      $ 2057 "Vial_liq_pick_3" "breakAfter"
      movel(Vial_liq_pick_3_p, a=0.5, v=0.1)
      $ 2058 "Vial_liq_pick_4" "breakAfter"
      movel(Vial_liq_pick_4_p, a=0.5, v=0.1)
      # begin: URCap Program Node
      #   Source: Robotiq_Grippers, 3.17.0.105337, Robotiq Inc.
      #   Type: Gripper
      $ 2059 "Gripper Close (1)"
      if not(gripper_connected[0]):
        popup("Gripper 1 must be connected to run this program.", "No connection", False, True, True)
      end
      if not(rq_is_gripper_activated("1")):
        popup("Gripper 1 is not activated. Go to Installation tab > Gripper to activate it and run the program again.", "Not activated", False, True, True)
      end
      rq_set_pos_spd_for(255, 82, 71, "1")
      rq_wait_pos_spe_for_request(255, 82, 71, "1")
      rq_go_to("1")
      rq_wait("1")
      # end: URCap Program Node
      $ 2060 "Wait: 1.0"
      sleep(1.0)
      $ 2061 "Set GRP_3F_Open=On"
      set_standard_digital_out(5, True)
      $ 2062 "Wait: 0.5"
      sleep(0.5)
      $ 2063 "Vial_liq_abov_2" "breakAfter"
      movel(Vial_liq_abov_2_p, a=0.3, v=0.05, r=0.05)
      $ 2064 "MoveL"
      $ 2065 "Liquid_midway_1" "breakAfter"
      movel(Liquid_midway_1_p, a=0.5, v=0.1)
      $ 2066 "Loop 3 times"
      Loop_1 = 0
      while (Loop_1 < 3):
        $ 2067 "shake_3" "breakAfter"
        movel(shake_3_p, a=2.0, v=0.5)
        $ 2068 "shake_4" "breakAfter"
        movel(shake_4_p, a=2.0, v=0.5)
        Loop_1 = Loop_1 + 1
      end
      $ 2069 "drop_above_3" "breakAfter"
      movel(drop_above_3_p, a=0.5, v=0.1)
      $ 2070 "drop_above_4" "breakAfter"
      movel(drop_above_4_p, a=0.5, v=0.1)
      $ 2071 "liq_tran_3" "breakAfter"
      movel(liq_tran_3_p, a=0.5, v=0.05, r=0.008)
      $ 2072 "Wait: 1.0"
      sleep(1.0)
      $ 2073 "drop_above_5" "breakAfter"
      movel(drop_above_5_p, a=0.5, v=0.1)
      $ 2074 "Waypoint_92" "breakAfter"
      movel(Waypoint_92_p, a=0.5, v=0.1)
      $ 2075 "liq_tran_4" "breakAfter"
      movel(liq_tran_4_p, a=0.5, v=0.05)
      $ 2076 "Wait: 1.0"
      sleep(1.0)
      $ 2077 "drop_above_6" "breakAfter"
      movel(drop_above_6_p, a=0.5, v=0.1)
      $ 2078 "drop_above_7" "breakAfter"
      movel(drop_above_7_p, a=0.5, v=0.1)
      $ 2079 "Liquid_midway_2" "breakAfter"
      movel(Liquid_midway_2_p, a=0.5, v=0.1)
      $ 2080 "MoveL"
      $ 2081 "Vial_drop_abo_1" "breakAfter"
      movel(Vial_drop_abo_1_p, a=0.5, v=0.1)
      $ 2082 "Vial_liq_drop_1" "breakAfter"
      movel(Vial_liq_drop_1_p, a=0.5, v=0.1)
      # begin: URCap Program Node
      #   Source: Robotiq_Grippers, 3.17.0.105337, Robotiq Inc.
      #   Type: Gripper
      $ 2083 "Gripper Open (1)"
      if not(gripper_connected[0]):
        popup("Gripper 1 must be connected to run this program.", "No connection", False, True, True)
      end
      if not(rq_is_gripper_activated("1")):
        popup("Gripper 1 is not activated. Go to Installation tab > Gripper to activate it and run the program again.", "Not activated", False, True, True)
      end
      rq_set_pos_spd_for(0, 82, 71, "1")
      rq_wait_pos_spe_for_request(0, 82, 71, "1")
      rq_go_to("1")
      rq_wait("1")
      # end: URCap Program Node
      $ 2084 "Vial_drop_abo_2" "breakAfter"
      movel(Vial_drop_abo_2_p, a=0.5, v=0.1)
    elif (34 == switch_1):
      $ 2085 "Case 34"
      $ 2086 "Task≔'Dosing'"
      global Task="Dosing"
      $ 2087 "tilt_to_home()"
      tilt_to_home()
      $ 2088 "Powder dosing all"
      $ 2089 "tilt_angle_sent≔0.0"
      global tilt_angle_sent=0.0
      $ 2090 "send_target_info()"
      send_target_info()
      $ 2092 "prev_spat≔''"
      global prev_spat=""
      $ 2093 "spatula≔''"
      global spatula=""
      $ 2094 "scoop_status≔'normal'"
      global scoop_status="normal"
      $ 2095 "send_powder_info()"
      send_powder_info()
      $ 2096 "Set AO[0]=0.0"
      set_standard_analog_out(0, 0.0)
      $ 2097 "Wait: 0.2"
      sleep(0.2)
      $ 2098 "reach pots decapping pose"
      # begin: URCap Program Node
      #   Source: SensoPart VISOR Robotic, 2.0.6, SensoPart Industriesensorik GmbH
      #   Type: VISOR Robotic App
      $ 2104 "VISOR Easy Pick"
      def visorFuncEasyPick_14c2cb():
        # begin: URCap Program Node
        #   Source: SensoPart VISOR Robotic, 2.0.6, SensoPart Industriesensorik GmbH
        #   Type: Easy Pick Setup
        $ 2105 "# 1 Setup" "noBreak"
        local easyPickVisorId = 1
        local easyPickArmMounted = True
        local easyPickSetJob = True
        local easyPickJobName = "Weight_scale"
        local easyPickAtImgAcq = False
        local easyPickImgAcqPose = Trigger
        # end: URCap Program Node
        # begin: URCap Program Node
        #   Source: SensoPart VISOR Robotic, 2.0.6, SensoPart Industriesensorik GmbH
        #   Type: Process
        $ 2106 "Process" "noBreak"
        local easyPickObjTaken = False
        local easyPickTrigger = False
        local easyPickPoseIdx = 0
        local easyPickPose = p[0,0,0,0,0,0]
        def easyPickFuncTrigger(visorId, setJob, jobName, arm):
        if (setJob):
          visor_changeJob(visorId, jobName, 6000)
        end
        if (arm):
          visor_trigger(visorId, 6000, "arm")
        else:
          visor_trigger(visorId, 6000)
        end
        global easyPickParts_4=visor_partsFound(visorId)
        visor_easyPickUpdate(visorId, "parts", visor_partsFound(visorId))
        return visor_getPose3d(visorId, 0)
      end
      while (not easyPickObjTaken):
        easyPickTrigger = (easyPickCount_4 >= visor_partsFound(easyPickVisorId)) or (easyPickCount_4 > 9) or (not visor_easyPickCheckIdent("850a49", easyPickVisorId))
        if (easyPickTrigger):
          easyPickCount_4 = 0
        end
        easyPickPoseIdx = easyPickCount_4
        easyPickPose = visor_getPose3d(easyPickVisorId, easyPickPoseIdx)
        visor_easyPickUpdate(easyPickVisorId, "counter", easyPickPoseIdx)
        # begin: URCap Program Node
        #   Source: SensoPart VISOR Robotic, 2.0.6, SensoPart Industriesensorik GmbH
        #   Type: Image Acquisition Pose
        $ 2107 "Image Acquisition Pose" "noBreak"
        if (easyPickTrigger):
          if (not easyPickAtImgAcq):
            movej(pose_trans(easyPickImgAcqPose,p[0.0000,0.0000,-0.0000,0.0000,0.0000,0.0000]),a=1.3963,v=1.0472,t=0.000000,r=0.000000)
            easyPickAtImgAcq = True
          end
          easyPickPose = easyPickFuncTrigger(easyPickVisorId, easyPickSetJob, easyPickJobName, easyPickArmMounted)
        end
        # end: URCap Program Node
        # begin: URCap Program Node
        #   Source: SensoPart VISOR Robotic, 2.0.6, SensoPart Industriesensorik GmbH
        #   Type: Object Detected
        $ 2108 "Object Detected" "noBreak"
        if (visor_partsFound(easyPickVisorId) > 0):
          $ 2109 "Open Gripper" "noBreak"
          $ 2110 "weight_value≔get_weight()" "noBreak"
          global weight_value=get_weight()
          $ 2111 "Wait: 0.5" "noBreak"
          sleep(0.5)
          $ 2112 "diff≔target_weight-weight_value" "noBreak"
          global diff=target_weight-weight_value
          $ 2113 "compute_level_percent(W_now, weight_value)" "noBreak"
          compute_level_percent(W_now, weight_value)
          $ 2114 "send_level_info()" "noBreak"
          send_level_info()
          $ 2115 "spatula≔select_spatula(Flowability, level, diff, bulk_density, mouth_d)" "noBreak"
          global spatula=select_spatula(Flowability, level, diff, bulk_density, mouth_d)
          $ 2116 "Wait: 0.2" "noBreak"
          sleep(0.2)
          $ 2117 "send_spatula_info()" "noBreak"
          send_spatula_info()
          $ 2118 "Pick spatula" "noBreak"
          $ 2119 "If spatula ≟ 'spatula_L'" "noBreak"
          if (spatula  ==  "spatula_L"):
            $ 2120 "MoveJ" "noBreak"
            $ 2121 "Spatula_otw" "noBreak"
            movej(get_inverse_kin(Spatula_otw_p, qnear=Spatula_otw_q), a=1.3962634015954636, v=1.0471975511965976)
            $ 2122 "pick_spat_L_abv" "noBreak"
            movej(get_inverse_kin(pick_spat_L_abv_p, qnear=pick_spat_L_abv_q), a=1.3962634015954636, v=1.0471975511965976)
            $ 2123 "MoveL" "noBreak"
            $ 2124 "spat_L_pick" "noBreak"
            movel(spat_L_pick_p, a=1.2, v=0.25)
            # begin: URCap Program Node
            #   Source: Robotiq_Grippers, 3.17.0.105337, Robotiq Inc.
            #   Type: Gripper
            $ 2125 "Gripper Close (1)" "noBreak"
            if not(gripper_connected[0]):
              popup("Gripper 1 must be connected to run this program.", "No connection", False, True, True)
            end
            if not(rq_is_gripper_activated("1")):
              popup("Gripper 1 is not activated. Go to Installation tab > Gripper to activate it and run the program again.", "Not activated", False, True, True)
            end
            rq_set_pos_spd_for(255, 0, 77, "1")
            rq_wait_pos_spe_for_request(255, 0, 77, "1")
            rq_go_to("1")
            rq_wait("1")
            # end: URCap Program Node
            $ 2126 "spat_L_lift" "noBreak"
            movel(spat_L_lift_p, a=1.2, v=0.25, r=0.01)
            $ 2127 "spat_L_side" "noBreak"
            movel(spat_L_side_p, a=1.2, v=0.25, r=0.01)
            $ 2128 "spat_L_up" "noBreak"
            movel(spat_L_up_p, a=1.2, v=0.25, r=0.05)
            $ 2129 "MoveJ" "noBreak"
            $ 2130 "Spatula_otw" "noBreak"
            movej(get_inverse_kin(Spatula_otw_p, qnear=Spatula_otw_q), a=1.3962634015954636, v=1.0471975511965976)
          else:
            $ 2131 "ElseIf spatula ≟'spatula_M'" "noBreak"
            if (spatula  == "spatula_M"):
              $ 2132 "MoveJ" "noBreak"
              $ 2133 "Spatula_otw" "noBreak"
              movej(get_inverse_kin(Spatula_otw_p, qnear=Spatula_otw_q), a=1.3962634015954636, v=1.0471975511965976)
              $ 2134 "spat_M_up" "noBreak"
              movej(get_inverse_kin(spat_M_up_p, qnear=spat_M_up_q), a=1.3962634015954636, v=1.0471975511965976, r=0.05)
              $ 2135 "MoveL" "noBreak"
              $ 2136 "spat_M_pick" "noBreak"
              movel(spat_M_pick_p, a=1.2, v=0.25)
              # begin: URCap Program Node
              #   Source: Robotiq_Grippers, 3.17.0.105337, Robotiq Inc.
              #   Type: Gripper
              $ 2137 "Gripper Close (1)" "noBreak"
              if not(gripper_connected[0]):
                popup("Gripper 1 must be connected to run this program.", "No connection", False, True, True)
              end
              if not(rq_is_gripper_activated("1")):
                popup("Gripper 1 is not activated. Go to Installation tab > Gripper to activate it and run the program again.", "Not activated", False, True, True)
              end
              rq_set_pos_spd_for(255, 0, 77, "1")
              rq_wait_pos_spe_for_request(255, 0, 77, "1")
              rq_go_to("1")
              rq_wait("1")
              # end: URCap Program Node
              $ 2138 "spat_M_up" "noBreak"
              movel(spat_M_up_p, a=1.2, v=0.25, r=0.05)
              $ 2139 "Spatula_otw" "noBreak"
              movel(Spatula_otw_p, a=1.2, v=0.25)
              $ 2140 "switch_spat_M≔ False " "noBreak"
              global switch_spat_M=  False
            else:
              $ 2141 "ElseIf spatula≟'spatula_S'" "noBreak"
              if (spatula == "spatula_S"):
                $ 2142 "MoveJ" "noBreak"
                $ 2143 "Spatula_otw" "noBreak"
                movej(get_inverse_kin(Spatula_otw_p, qnear=Spatula_otw_q), a=1.3962634015954636, v=1.0471975511965976)
                $ 2144 "spat_S_Up_7" "noBreak"
                movej(get_inverse_kin(spat_S_Up_7_p, qnear=spat_S_Up_7_q), a=1.3962634015954636, v=1.0471975511965976, r=0.05)
                $ 2145 "MoveL" "noBreak"
                $ 2146 "spat_S_Pick_4" "noBreak"
                movel(spat_S_Pick_4_p, a=1.2, v=0.25)
                # begin: URCap Program Node
                #   Source: Robotiq_Grippers, 3.17.0.105337, Robotiq Inc.
                #   Type: Gripper
                $ 2147 "Gripper Close (1)" "noBreak"
                if not(gripper_connected[0]):
                  popup("Gripper 1 must be connected to run this program.", "No connection", False, True, True)
                end
                if not(rq_is_gripper_activated("1")):
                  popup("Gripper 1 is not activated. Go to Installation tab > Gripper to activate it and run the program again.", "Not activated", False, True, True)
                end
                rq_set_pos_spd_for(255, 0, 77, "1")
                rq_wait_pos_spe_for_request(255, 0, 77, "1")
                rq_go_to("1")
                rq_wait("1")
                # end: URCap Program Node
                $ 2148 "spat_S_Up_8" "noBreak"
                movel(spat_S_Up_8_p, a=1.2, v=0.25, r=0.05)
                $ 2149 "Spatula_otw" "noBreak"
                movel(Spatula_otw_p, a=1.2, v=0.25)
                $ 2150 "switch_spat_S≔ False " "noBreak"
                global switch_spat_S=  False
              else:
                $ 2151 "ElseIf spatula≟'spatula_flat_M'" "noBreak"
                if (spatula == "spatula_flat_M"):
                  $ 2152 "MoveJ" "noBreak"
                  $ 2153 "Spatula_otw" "noBreak"
                  movej(get_inverse_kin(Spatula_otw_p, qnear=Spatula_otw_q), a=1.3962634015954636, v=1.0471975511965976)
                  $ 2154 "spat_flatM_up" "noBreak"
                  movej(get_inverse_kin(spat_flatM_up_p, qnear=spat_flatM_up_q), a=1.3962634015954636, v=1.0471975511965976, r=0.05)
                  $ 2155 "MoveL" "noBreak"
                  $ 2156 "spat_flatM_pick" "noBreak"
                  movel(spat_flatM_pick_p, a=1.2, v=0.25)
                  # begin: URCap Program Node
                  #   Source: Robotiq_Grippers, 3.17.0.105337, Robotiq Inc.
                  #   Type: Gripper
                  $ 2157 "Gripper Close (1)" "noBreak"
                  if not(gripper_connected[0]):
                    popup("Gripper 1 must be connected to run this program.", "No connection", False, True, True)
                  end
                  if not(rq_is_gripper_activated("1")):
                    popup("Gripper 1 is not activated. Go to Installation tab > Gripper to activate it and run the program again.", "Not activated", False, True, True)
                  end
                  rq_set_pos_spd_for(255, 0, 77, "1")
                  rq_wait_pos_spe_for_request(255, 0, 77, "1")
                  rq_go_to("1")
                  rq_wait("1")
                  # end: URCap Program Node
                  $ 2158 "spat_flatM_up" "noBreak"
                  movel(spat_flatM_up_p, a=1.2, v=0.25, r=0.05)
                  $ 2159 "Spatula_otw" "noBreak"
                  movel(Spatula_otw_p, a=1.2, v=0.25)
                  $ 2160 "switch_spat_F_M≔ False " "noBreak"
                  global switch_spat_F_M=  False
                else:
                  $ 2161 "ElseIf spatula≟'spatula_flat_S'" "noBreak"
                  if (spatula == "spatula_flat_S"):
                    $ 2162 "MoveJ" "noBreak"
                    $ 2163 "Spatula_otw" "noBreak"
                    movej(get_inverse_kin(Spatula_otw_p, qnear=Spatula_otw_q), a=1.3962634015954636, v=1.0471975511965976)
                    $ 2164 "spat_flatS_up" "noBreak"
                    movej(get_inverse_kin(spat_flatS_up_p, qnear=spat_flatS_up_q), a=1.3962634015954636, v=1.0471975511965976, r=0.05)
                    $ 2165 "MoveL" "noBreak"
                    $ 2166 "spat_flatS_pick" "noBreak"
                    movel(spat_flatS_pick_p, a=1.2, v=0.25)
                    # begin: URCap Program Node
                    #   Source: Robotiq_Grippers, 3.17.0.105337, Robotiq Inc.
                    #   Type: Gripper
                    $ 2167 "Gripper Close (1)" "noBreak"
                    if not(gripper_connected[0]):
                      popup("Gripper 1 must be connected to run this program.", "No connection", False, True, True)
                    end
                    if not(rq_is_gripper_activated("1")):
                      popup("Gripper 1 is not activated. Go to Installation tab > Gripper to activate it and run the program again.", "Not activated", False, True, True)
                    end
                    rq_set_pos_spd_for(255, 0, 77, "1")
                    rq_wait_pos_spe_for_request(255, 0, 77, "1")
                    rq_go_to("1")
                    rq_wait("1")
                    # end: URCap Program Node
                    $ 2168 "spat_flatS_up" "noBreak"
                    movel(spat_flatS_up_p, a=1.2, v=0.25, r=0.05)
                    $ 2169 "Spatula_otw" "noBreak"
                    movel(Spatula_otw_p, a=1.2, v=0.25)
                    $ 2170 "switch_spat_F_S≔ False " "noBreak"
                    global switch_spat_F_S=  False
                  end
                end
              end
            end
          end
          $ 2171 "Action_Info≔'Scooping'" "noBreak"
          global Action_Info="Scooping"
          $ 2172 "auto_tilt_and_scoop(W_now, target_weight, weight_value)" "noBreak"
          auto_tilt_and_scoop(W_now, target_weight, weight_value)
          $ 2173 "Action_Info≔'Dosing'" "noBreak"
          global Action_Info="Dosing"
          # begin: URCap Program Node
          #   Source: SensoPart VISOR Robotic, 2.0.6, SensoPart Industriesensorik GmbH
          #   Type: Approach Pose
          $ 2174 "Approach Pose" "noBreak"
          movej(pose_trans(easyPickPose,p[0.0000,0.0000,-0.0000,0.0000,0.0000,0.0000]),a=0.2618,v=0.1745,t=0.000000,r=0.000000)
          # end: URCap Program Node
          # begin: URCap Program Node
          #   Source: SensoPart VISOR Robotic, 2.0.6, SensoPart Industriesensorik GmbH
          #   Type: Target Pose
          $ 2175 "Target Pose" "noBreak"
          movel(pose_trans(easyPickPose,p[0.0000,0.0000,-0.0000,0.0000,0.0000,0.0000]),a=0.0500,v=0.0200,t=0.000000,r=0.000000)
          # end: URCap Program Node
          $ 2176 "Close Gripper" "noBreak"
          $ 2177 "current_p≔get_actual_tcp_pose()" "noBreak"
          global current_p= get_actual_tcp_pose ()
          $ 2178 "dispense_pos≔pose_trans(current_p,p[0,0,0,0,-deg2rad(spatula_ry),0])" "noBreak"
          global dispense_pos=pose_trans(current_p,p[0,0,0,0,-deg2rad(spatula_ry),0])
          $ 2180 "Loop weight_value≤target_weight " "noBreak"
          thread Thread_while_2180():
            while (True):
              $ 2181 "MoveL" "noBreak"
              $ 2182 "dispense_pos" "noBreak"
              movel(dispense_pos, a=0.2, v=0.1)
              $ 2183 "log_weight()" "noBreak"
              log_weight()
              $ 2185 "CCW_full_Rotate()" "noBreak"
              CCW_full_Rotate()
              $ 2186 "Start_thread≔ True " "noBreak"
              global Start_thread=  True
              $ 2187 "vib_thread≔ True " "noBreak"
              global vib_thread=  True
              $ 2188 "Wait: 0.5" "noBreak"
              sleep(0.5)
              $ 2189 "If diff ≥(target_g*1.2)" "noBreak"
              if (diff  >= (target_g*1.2)):
                $ 2190 "tilt_pose≔pose_trans(get_actual_tcp_pose(), p[0, 0, 0, 0, 0, 2.0])" "noBreak"
                global tilt_pose=pose_trans(get_actual_tcp_pose(), p[0, 0, 0, 0, 0, 2.0])
                $ 2191 "movel(tilt_pose, a=0.5, v=0.5, r=0.00001)" "noBreak"
                movel(tilt_pose, a=0.5, v=0.5, r=0.00001)
              else:
                $ 2192 "Else" "noBreak"
                $ 2193 "Loop weight_value≤(target_weight-0.00) and tilt_angle≥(-1.999) and tilt_angle≤0.5" "noBreak"
                thread Thread_while_2193():
                  while (True):
                    $ 2194 "current_error≔target_weight-weight_value" "noBreak"
                    global current_error=target_weight-weight_value
                    $ 2195 "Integral_error≔Integral_error+current_error*dt" "noBreak"
                    global Integral_error=Integral_error+current_error*dt
                    $ 2196 "derivative≔(current_error-previous_error)/dt" "noBreak"
                    global derivative=(current_error-previous_error)/dt
                    $ 2197 "tilt_increment≔(kp*current_error)+(ki*Integral_error)+(kd*derivative)" "noBreak"
                    global tilt_increment=(kp*current_error)+(ki*Integral_error)+(kd*derivative)
                    $ 2198 "current_pose≔get_actual_tcp_pose()" "noBreak"
                    global current_pose= get_actual_tcp_pose ()
                    $ 2199 "tilt_angle≔current_pose[5]" "noBreak"
                    global tilt_angle=current_pose[5]
                    $ 2200 "tilt_pose≔pose_trans(current_pose, p[0, 0, 0, 0, 0, tilt_increment])" "noBreak"
                    global tilt_pose=pose_trans(current_pose, p[0, 0, 0, 0, 0, tilt_increment])
                    $ 2201 "movel(tilt_pose, a=0.1, v=0.1, r=0.00001)" "noBreak"
                    movel(tilt_pose, a=0.1, v=0.1, r=0.00001)
                    $ 2202 "previous_error≔current_error" "noBreak"
                    global previous_error=current_error
                  end
                end
                if (weight_value <= (target_weight-0.00)  and  tilt_angle >= (-1.999)  and  tilt_angle <= 0.5):
                  global thread_handler_2193=run Thread_while_2193()
                  while (weight_value <= (target_weight-0.00)  and  tilt_angle >= (-1.999)  and  tilt_angle <= 0.5):
                    sync()
                  end
                  kill thread_handler_2193
                end
              end
              $ 2203 "weight_value≔get_weight()" "noBreak"
              global weight_value=get_weight()
              $ 2205 "tilt_angle≔-1" "noBreak"
              global tilt_angle=-1
              $ 2206 "Wait: 0.5" "noBreak"
              sleep(0.5)
              $ 2207 "Start_thread≔ False " "noBreak"
              global Start_thread=  False
              $ 2208 "vib_thread≔ False " "noBreak"
              global vib_thread=  False
              $ 2210 "dispense_pos" "noBreak"
              movel(dispense_pos, a=1.2, v=0.25)
              $ 2211 "compute_level_percent(W_now, weight_value)" "noBreak"
              compute_level_percent(W_now, weight_value)
              $ 2212 "prev_spat≔spatula" "noBreak"
              global prev_spat=spatula
              $ 2213 "Wait: 0.2" "noBreak"
              sleep(0.2)
              $ 2214 "spatula≔select_spatula(Flowability, level, diff, bulk_density, mouth_d)" "noBreak"
              global spatula=select_spatula(Flowability, level, diff, bulk_density, mouth_d)
              $ 2215 "Wait: 1.0" "noBreak"
              sleep(1.0)
              $ 2216 "send_level_info()" "noBreak"
              send_level_info()
              $ 2217 "send_spatula_info()" "noBreak"
              send_spatula_info()
              $ 2218 "Integral_error≔0" "noBreak"
              global Integral_error=0
              $ 2219 "current_error≔0" "noBreak"
              global current_error=0
              $ 2220 "previous_error≔0" "noBreak"
              global previous_error=0
              $ 2221 "Set AO[0]=0.0" "noBreak"
              set_standard_analog_out(0, 0.0)
              $ 2222 "Wait: 0.5" "noBreak"
              sleep(0.5)
              $ 2223 "swtich spatula" "noBreak"
              $ 2224 "If spatula ≟ 'spatula_M' and switch_spat_M≟ True " "noBreak"
              if (spatula  ==  "spatula_M"  and  switch_spat_M ==   True  ):
                $ 2225 "MoveJ" "noBreak"
                $ 2226 "Spatula_otw" "noBreak"
                movej(get_inverse_kin(Spatula_otw_p, qnear=Spatula_otw_q), a=1.3962634015954636, v=1.0471975511965976)
                $ 2227 "spat_L_up" "noBreak"
                movej(get_inverse_kin(spat_L_up_p, qnear=spat_L_up_q), a=1.3962634015954636, v=1.0471975511965976)
                $ 2228 "MoveL" "noBreak"
                $ 2229 "spat_L_side" "noBreak"
                movel(spat_L_side_p, a=1.2, v=0.25)
                $ 2230 "spat_L_lift" "noBreak"
                movel(spat_L_lift_p, a=1.2, v=0.25)
                $ 2231 "spat_L_pick" "noBreak"
                movel(spat_L_pick_p, a=0.2, v=0.1)
                # begin: URCap Program Node
                #   Source: Robotiq_Grippers, 3.17.0.105337, Robotiq Inc.
                #   Type: Gripper
                $ 2232 "Gripper Open (1)" "noBreak"
                if not(gripper_connected[0]):
                  popup("Gripper 1 must be connected to run this program.", "No connection", False, True, True)
                end
                if not(rq_is_gripper_activated("1")):
                  popup("Gripper 1 is not activated. Go to Installation tab > Gripper to activate it and run the program again.", "Not activated", False, True, True)
                end
                rq_set_pos_spd_for(0, 255, 77, "1")
                rq_wait_pos_spe_for_request(0, 255, 77, "1")
                rq_go_to("1")
                rq_wait("1")
                # end: URCap Program Node
                $ 2233 "spat_M_pick" "noBreak"
                movel(spat_M_pick_p, a=1.2, v=0.25)
                # begin: URCap Program Node
                #   Source: Robotiq_Grippers, 3.17.0.105337, Robotiq Inc.
                #   Type: Gripper
                $ 2234 "Gripper Close (1)" "noBreak"
                if not(gripper_connected[0]):
                  popup("Gripper 1 must be connected to run this program.", "No connection", False, True, True)
                end
                if not(rq_is_gripper_activated("1")):
                  popup("Gripper 1 is not activated. Go to Installation tab > Gripper to activate it and run the program again.", "Not activated", False, True, True)
                end
                rq_set_pos_spd_for(255, 0, 77, "1")
                rq_wait_pos_spe_for_request(255, 0, 77, "1")
                rq_go_to("1")
                rq_wait("1")
                # end: URCap Program Node
                $ 2235 "spat_M_up" "noBreak"
                movel(spat_M_up_p, a=1.2, v=0.25)
                $ 2236 "Spatula_otw" "noBreak"
                movel(Spatula_otw_p, a=1.2, v=0.25)
                $ 2237 "switch_spat_M≔ False " "noBreak"
                global switch_spat_M=  False
                $ 2238 "correction_reset()" "noBreak"
                correction_reset()
              else:
                $ 2239 "ElseIf spatula ≟ 'spatula_S' and switch_spat_S ≟ True and prev_spat≟'spatula_M'" "noBreak"
                if (spatula  ==  "spatula_S" and switch_spat_S  ==   True  and prev_spat == "spatula_M"):
                  $ 2240 "MoveL" "noBreak"
                  $ 2241 "Spatula_otw" "noBreak"
                  movel(Spatula_otw_p, a=1.2, v=0.25)
                  $ 2242 "spat_M_up" "noBreak"
                  movel(spat_M_up_p, a=1.2, v=0.25)
                  $ 2243 "spat_M_pick" "noBreak"
                  movel(spat_M_pick_p, a=0.2, v=0.1)
                  # begin: URCap Program Node
                  #   Source: Robotiq_Grippers, 3.17.0.105337, Robotiq Inc.
                  #   Type: Gripper
                  $ 2244 "Gripper Open (1)" "noBreak"
                  if not(gripper_connected[0]):
                    popup("Gripper 1 must be connected to run this program.", "No connection", False, True, True)
                  end
                  if not(rq_is_gripper_activated("1")):
                    popup("Gripper 1 is not activated. Go to Installation tab > Gripper to activate it and run the program again.", "Not activated", False, True, True)
                  end
                  rq_set_pos_spd_for(0, 255, 77, "1")
                  rq_wait_pos_spe_for_request(0, 255, 77, "1")
                  rq_go_to("1")
                  rq_wait("1")
                  # end: URCap Program Node
                  $ 2245 "spat_S_pick" "noBreak"
                  movel(spat_S_pick_p, a=1.2, v=0.25)
                  # begin: URCap Program Node
                  #   Source: Robotiq_Grippers, 3.17.0.105337, Robotiq Inc.
                  #   Type: Gripper
                  $ 2246 "Gripper Close (1)" "noBreak"
                  if not(gripper_connected[0]):
                    popup("Gripper 1 must be connected to run this program.", "No connection", False, True, True)
                  end
                  if not(rq_is_gripper_activated("1")):
                    popup("Gripper 1 is not activated. Go to Installation tab > Gripper to activate it and run the program again.", "Not activated", False, True, True)
                  end
                  rq_set_pos_spd_for(255, 0, 77, "1")
                  rq_wait_pos_spe_for_request(255, 0, 77, "1")
                  rq_go_to("1")
                  rq_wait("1")
                  # end: URCap Program Node
                  $ 2247 "spat_S_up" "noBreak"
                  movel(spat_S_up_p, a=1.2, v=0.25)
                  $ 2248 "Spatula_otw" "noBreak"
                  movel(Spatula_otw_p, a=1.2, v=0.25)
                  $ 2249 "switch_spat_S≔ False " "noBreak"
                  global switch_spat_S=  False
                  $ 2250 "correction_reset()" "noBreak"
                  correction_reset()
                else:
                  $ 2251 "ElseIf spatula≟'spatula_S' and switch_spat_S≟ True  and prev_spat≟'spatula_L'" "noBreak"
                  if (spatula == "spatula_S" and switch_spat_S ==   True    and  prev_spat == "spatula_L"):
                    $ 2252 "MoveJ" "noBreak"
                    $ 2253 "Spatula_otw" "noBreak"
                    movej(get_inverse_kin(Spatula_otw_p, qnear=Spatula_otw_q), a=1.3962634015954636, v=1.0471975511965976)
                    $ 2254 "spat_L_up" "noBreak"
                    movej(get_inverse_kin(spat_L_up_p, qnear=spat_L_up_q), a=1.3962634015954636, v=1.0471975511965976)
                    $ 2255 "MoveL" "noBreak"
                    $ 2256 "spat_L_side" "noBreak"
                    movel(spat_L_side_p, a=1.2, v=0.25)
                    $ 2257 "spat_L_lift" "noBreak"
                    movel(spat_L_lift_p, a=1.2, v=0.25)
                    $ 2258 "spat_L_pick" "noBreak"
                    movel(spat_L_pick_p, a=0.2, v=0.1)
                    # begin: URCap Program Node
                    #   Source: Robotiq_Grippers, 3.17.0.105337, Robotiq Inc.
                    #   Type: Gripper
                    $ 2259 "Gripper Open (1)" "noBreak"
                    if not(gripper_connected[0]):
                      popup("Gripper 1 must be connected to run this program.", "No connection", False, True, True)
                    end
                    if not(rq_is_gripper_activated("1")):
                      popup("Gripper 1 is not activated. Go to Installation tab > Gripper to activate it and run the program again.", "Not activated", False, True, True)
                    end
                    rq_set_pos_spd_for(0, 255, 77, "1")
                    rq_wait_pos_spe_for_request(0, 255, 77, "1")
                    rq_go_to("1")
                    rq_wait("1")
                    # end: URCap Program Node
                    $ 2260 "spat_S_pick" "noBreak"
                    movel(spat_S_pick_p, a=1.2, v=0.25)
                    # begin: URCap Program Node
                    #   Source: Robotiq_Grippers, 3.17.0.105337, Robotiq Inc.
                    #   Type: Gripper
                    $ 2261 "Gripper Close (1)" "noBreak"
                    if not(gripper_connected[0]):
                      popup("Gripper 1 must be connected to run this program.", "No connection", False, True, True)
                    end
                    if not(rq_is_gripper_activated("1")):
                      popup("Gripper 1 is not activated. Go to Installation tab > Gripper to activate it and run the program again.", "Not activated", False, True, True)
                    end
                    rq_set_pos_spd_for(255, 0, 77, "1")
                    rq_wait_pos_spe_for_request(255, 0, 77, "1")
                    rq_go_to("1")
                    rq_wait("1")
                    # end: URCap Program Node
                    $ 2262 "spat_S_up" "noBreak"
                    movel(spat_S_up_p, a=1.2, v=0.25)
                    $ 2263 "Spatula_otw" "noBreak"
                    movel(Spatula_otw_p, a=1.2, v=0.25)
                    $ 2264 "switch_spat_S≔ False " "noBreak"
                    global switch_spat_S=  False
                    $ 2265 "correction_reset()" "noBreak"
                    correction_reset()
                  else:
                    $ 2266 "ElseIf spatula≟'spatula_flat_S'  and switch_spat_F_S ≟ True " "noBreak"
                    if (spatula == "spatula_flat_S"   and  switch_spat_F_S  ==   True  ):
                      $ 2267 "MoveL" "noBreak"
                      $ 2268 "Spatula_otw" "noBreak"
                      movel(Spatula_otw_p, a=1.2, v=0.25)
                      $ 2269 "spat_flatM_up" "noBreak"
                      movel(spat_flatM_up_p, a=1.2, v=0.25)
                      $ 2270 "spat_flatM_pick" "noBreak"
                      movel(spat_flatM_pick_p, a=0.2, v=0.1)
                      # begin: URCap Program Node
                      #   Source: Robotiq_Grippers, 3.17.0.105337, Robotiq Inc.
                      #   Type: Gripper
                      $ 2271 "Gripper Open (1)" "noBreak"
                      if not(gripper_connected[0]):
                        popup("Gripper 1 must be connected to run this program.", "No connection", False, True, True)
                      end
                      if not(rq_is_gripper_activated("1")):
                        popup("Gripper 1 is not activated. Go to Installation tab > Gripper to activate it and run the program again.", "Not activated", False, True, True)
                      end
                      rq_set_pos_spd_for(0, 255, 74, "1")
                      rq_wait_pos_spe_for_request(0, 255, 74, "1")
                      rq_go_to("1")
                      rq_wait("1")
                      # end: URCap Program Node
                      $ 2272 "spat_flatS_pick" "noBreak"
                      movel(spat_flatS_pick_p, a=1.2, v=0.25)
                      # begin: URCap Program Node
                      #   Source: Robotiq_Grippers, 3.17.0.105337, Robotiq Inc.
                      #   Type: Gripper
                      $ 2273 "Gripper Close (1)" "noBreak"
                      if not(gripper_connected[0]):
                        popup("Gripper 1 must be connected to run this program.", "No connection", False, True, True)
                      end
                      if not(rq_is_gripper_activated("1")):
                        popup("Gripper 1 is not activated. Go to Installation tab > Gripper to activate it and run the program again.", "Not activated", False, True, True)
                      end
                      rq_set_pos_spd_for(255, 0, 77, "1")
                      rq_wait_pos_spe_for_request(255, 0, 77, "1")
                      rq_go_to("1")
                      rq_wait("1")
                      # end: URCap Program Node
                      $ 2274 "spat_flatS_up" "noBreak"
                      movel(spat_flatS_up_p, a=1.2, v=0.25)
                      $ 2275 "Spatula_otw" "noBreak"
                      movel(Spatula_otw_p, a=1.2, v=0.25)
                      $ 2276 "switch_spat_F_S≔ False " "noBreak"
                      global switch_spat_F_S=  False
                      $ 2277 "correction_reset()" "noBreak"
                      correction_reset()
                    end
                  end
                end
              end
              $ 2278 "tilt(level)" "noBreak"
              tilt(level)
              $ 2279 "Action_Info≔'Scooping'" "noBreak"
              global Action_Info="Scooping"
              $ 2280 "auto_tilt_and_scoop(W_now, target_weight, weight_value)" "noBreak"
              auto_tilt_and_scoop(W_now, target_weight, weight_value)
              $ 2281 "Action_Info≔'Dosing'" "noBreak"
              global Action_Info="Dosing"
            end
          end
          if (weight_value <= target_weight ):
            global thread_handler_2180=run Thread_while_2180()
            while (weight_value <= target_weight ):
              sync()
            end
            kill thread_handler_2180
          end
          $ 2282 "Start_thread≔ False " "noBreak"
          global Start_thread=  False
          $ 2283 "vib_thread≔ False " "noBreak"
          global vib_thread=  False
          # begin: URCap Program Node
          #   Source: SensoPart VISOR Robotic, 2.0.6, SensoPart Industriesensorik GmbH
          #   Type: Exit Pose
          $ 2284 "Exit Pose" "noBreak"
          movel(pose_trans(easyPickPose,p[0.0000,0.0000,-0.0000,0.0000,0.0000,0.0000]),a=0.5000,v=0.2500,t=0.000000,r=0.000000)
          # end: URCap Program Node
          easyPickObjTaken = True
        end
        # end: URCap Program Node
        # begin: URCap Program Node
        #   Source: SensoPart VISOR Robotic, 2.0.6, SensoPart Industriesensorik GmbH
        #   Type: No Object Detected
        $ 2285 "No Object Detected" "noBreak"
        if (visor_partsFound(easyPickVisorId) < 1):
          $ 2286 "Popup: No weigh scale detected" "noBreak"
          popup("No weigh scale detected", "Message", False, False, blocking=True)
          else:
        end
        # end: URCap Program Node
      end
      easyPickCount_4 = easyPickCount_4 + 1
      visor_easyPickUpdate(easyPickVisorId, "counter", easyPickCount_4)
      visor_easyPickSetIdent("850a49", easyPickVisorId)
      # end: URCap Program Node
    end
    visorFuncEasyPick_14c2cb()
    # end: URCap Program Node
    $ 2287 "MoveL"
    $ 2288 "dispense_pos" "breakAfter"
    movel(dispense_pos, a=0.2, v=0.1)
    $ 2289 "after_scoop()"
    after_scoop()
    $ 2290 "Place spatula back to the rack"
    $ 2291 "If spatula ≟ 'spatula_L'"
    if (spatula  ==  "spatula_L"):
      $ 2292 "MoveJ"
      $ 2293 "Spatula_otw" "breakAfter"
      movej(get_inverse_kin(Spatula_otw_p, qnear=Spatula_otw_q), a=1.3962634015954636, v=1.0471975511965976)
      $ 2294 "MoveL"
      $ 2295 "spat_L_up" "breakAfter"
      movel(spat_L_up_p, a=1.2, v=0.25, r=0.05)
      $ 2296 "spat_L_side" "breakAfter"
      movel(spat_L_side_p, a=1.2, v=0.25, r=0.01)
      $ 2297 "spat_L_lift" "breakAfter"
      movel(spat_L_lift_p, a=1.2, v=0.25, r=0.01)
      $ 2298 "spat_L_pick" "breakAfter"
      movel(spat_L_pick_p, a=0.2, v=0.1)
      # begin: URCap Program Node
      #   Source: Robotiq_Grippers, 3.17.0.105337, Robotiq Inc.
      #   Type: Gripper
      $ 2299 "Gripper Open (1)"
      if not(gripper_connected[0]):
        popup("Gripper 1 must be connected to run this program.", "No connection", False, True, True)
      end
      if not(rq_is_gripper_activated("1")):
        popup("Gripper 1 is not activated. Go to Installation tab > Gripper to activate it and run the program again.", "Not activated", False, True, True)
      end
      rq_set_pos_spd_for(0, 128, 128, "1")
      rq_wait_pos_spe_for_request(0, 128, 128, "1")
      rq_go_to("1")
      rq_wait("1")
      # end: URCap Program Node
      $ 2300 "MoveJ"
      $ 2301 "pick_spat_L_abv" "breakAfter"
      movej(get_inverse_kin(pick_spat_L_abv_p, qnear=pick_spat_L_abv_q), a=1.3962634015954636, v=1.0471975511965976)
      $ 2302 "Spatula_otw" "breakAfter"
      movej(get_inverse_kin(Spatula_otw_p, qnear=Spatula_otw_q), a=1.3962634015954636, v=1.0471975511965976)
    else:
      $ 2303 "ElseIf spatula ≟'spatula_M'"
      if (spatula  == "spatula_M"):
        $ 2304 "MoveJ"
        $ 2305 "Spatula_otw" "breakAfter"
        movej(get_inverse_kin(Spatula_otw_p, qnear=Spatula_otw_q), a=1.3962634015954636, v=1.0471975511965976)
        $ 2306 "spat_M_up" "breakAfter"
        movej(get_inverse_kin(spat_M_up_p, qnear=spat_M_up_q), a=1.3962634015954636, v=1.0471975511965976, r=0.05)
        $ 2307 "MoveL"
        $ 2308 "spat_M_pick" "breakAfter"
        movel(spat_M_pick_p, a=0.2, v=0.1)
        # begin: URCap Program Node
        #   Source: Robotiq_Grippers, 3.17.0.105337, Robotiq Inc.
        #   Type: Gripper
        $ 2309 "Gripper Open (1)"
        if not(gripper_connected[0]):
          popup("Gripper 1 must be connected to run this program.", "No connection", False, True, True)
        end
        if not(rq_is_gripper_activated("1")):
          popup("Gripper 1 is not activated. Go to Installation tab > Gripper to activate it and run the program again.", "Not activated", False, True, True)
        end
        rq_set_pos_spd_for(0, 128, 128, "1")
        rq_wait_pos_spe_for_request(0, 128, 128, "1")
        rq_go_to("1")
        rq_wait("1")
        # end: URCap Program Node
        $ 2310 "spat_M_up" "breakAfter"
        movel(spat_M_up_p, a=1.2, v=0.25, r=0.05)
        $ 2311 "Spatula_otw" "breakAfter"
        movel(Spatula_otw_p, a=1.2, v=0.25)
        $ 2312 "switch_spat_M≔ False "
        global switch_spat_M=  False
      else:
        $ 2313 "ElseIf spatula≟'spatula_S'"
        if (spatula == "spatula_S"):
          $ 2314 "MoveJ"
          $ 2315 "Spatula_otw" "breakAfter"
          movej(get_inverse_kin(Spatula_otw_p, qnear=Spatula_otw_q), a=1.3962634015954636, v=1.0471975511965976)
          $ 2316 "spat_S_Up_7" "breakAfter"
          movej(get_inverse_kin(spat_S_Up_7_p, qnear=spat_S_Up_7_q), a=1.3962634015954636, v=1.0471975511965976, r=0.05)
          $ 2317 "MoveL"
          $ 2318 "spat_S_Pick_4" "breakAfter"
          movel(spat_S_Pick_4_p, a=0.2, v=0.1)
          # begin: URCap Program Node
          #   Source: Robotiq_Grippers, 3.17.0.105337, Robotiq Inc.
          #   Type: Gripper
          $ 2319 "Gripper Open (1)"
          if not(gripper_connected[0]):
            popup("Gripper 1 must be connected to run this program.", "No connection", False, True, True)
          end
          if not(rq_is_gripper_activated("1")):
            popup("Gripper 1 is not activated. Go to Installation tab > Gripper to activate it and run the program again.", "Not activated", False, True, True)
          end
          rq_set_pos_spd_for(0, 255, 51, "1")
          rq_wait_pos_spe_for_request(0, 255, 51, "1")
          rq_go_to("1")
          rq_wait("1")
          # end: URCap Program Node
          $ 2320 "spat_S_Up_8" "breakAfter"
          movel(spat_S_Up_8_p, a=1.2, v=0.25, r=0.05)
          $ 2321 "Spatula_otw" "breakAfter"
          movel(Spatula_otw_p, a=1.2, v=0.25)
          $ 2322 "switch_spat_S≔ False "
          global switch_spat_S=  False
        else:
          $ 2323 "ElseIf spatula≟'spatula_flat_M'"
          if (spatula == "spatula_flat_M"):
            $ 2324 "MoveJ"
            $ 2325 "Spatula_otw" "breakAfter"
            movej(get_inverse_kin(Spatula_otw_p, qnear=Spatula_otw_q), a=1.3962634015954636, v=1.0471975511965976)
            $ 2326 "spat_flatM_up" "breakAfter"
            movej(get_inverse_kin(spat_flatM_up_p, qnear=spat_flatM_up_q), a=1.3962634015954636, v=1.0471975511965976, r=0.05)
            $ 2327 "MoveL"
            $ 2328 "spat_flatM_pick" "breakAfter"
            movel(spat_flatM_pick_p, a=0.2, v=0.1)
            # begin: URCap Program Node
            #   Source: Robotiq_Grippers, 3.17.0.105337, Robotiq Inc.
            #   Type: Gripper
            $ 2329 "Gripper Open (1)"
            if not(gripper_connected[0]):
              popup("Gripper 1 must be connected to run this program.", "No connection", False, True, True)
            end
            if not(rq_is_gripper_activated("1")):
              popup("Gripper 1 is not activated. Go to Installation tab > Gripper to activate it and run the program again.", "Not activated", False, True, True)
            end
            rq_set_pos_spd_for(0, 128, 128, "1")
            rq_wait_pos_spe_for_request(0, 128, 128, "1")
            rq_go_to("1")
            rq_wait("1")
            # end: URCap Program Node
            $ 2330 "spat_flatM_up" "breakAfter"
            movel(spat_flatM_up_p, a=1.2, v=0.25, r=0.05)
            $ 2331 "Spatula_otw" "breakAfter"
            movel(Spatula_otw_p, a=1.2, v=0.25)
            $ 2332 "switch_spat_F_M≔ False "
            global switch_spat_F_M=  False
          else:
            $ 2333 "ElseIf spatula≟'spatula_flat_S'"
            if (spatula == "spatula_flat_S"):
              $ 2334 "MoveJ"
              $ 2335 "Spatula_otw" "breakAfter"
              movej(get_inverse_kin(Spatula_otw_p, qnear=Spatula_otw_q), a=1.3962634015954636, v=1.0471975511965976)
              $ 2336 "spat_flatS_up" "breakAfter"
              movej(get_inverse_kin(spat_flatS_up_p, qnear=spat_flatS_up_q), a=1.3962634015954636, v=1.0471975511965976, r=0.05)
              $ 2337 "MoveL"
              $ 2338 "spat_flatS_pick" "breakAfter"
              movel(spat_flatS_pick_p, a=0.2, v=0.1)
              # begin: URCap Program Node
              #   Source: Robotiq_Grippers, 3.17.0.105337, Robotiq Inc.
              #   Type: Gripper
              $ 2339 "Gripper Open (1)"
              if not(gripper_connected[0]):
                popup("Gripper 1 must be connected to run this program.", "No connection", False, True, True)
              end
              if not(rq_is_gripper_activated("1")):
                popup("Gripper 1 is not activated. Go to Installation tab > Gripper to activate it and run the program again.", "Not activated", False, True, True)
              end
              rq_set_pos_spd_for(0, 128, 128, "1")
              rq_wait_pos_spe_for_request(0, 128, 128, "1")
              rq_go_to("1")
              rq_wait("1")
              # end: URCap Program Node
              $ 2340 "spat_flatS_up" "breakAfter"
              movel(spat_flatS_up_p, a=1.2, v=0.25, r=0.05)
              $ 2341 "Spatula_otw" "breakAfter"
              movel(Spatula_otw_p, a=1.2, v=0.25)
              $ 2342 "switch_spat_F_S≔ False "
              global switch_spat_F_S=  False
            end
          end
        end
      end
    end
    $ 2343 "switch_spat_M≔ True "
    global switch_spat_M=  True
    $ 2344 "switch_spat_S≔ True "
    global switch_spat_S=  True
    $ 2345 "switch_spat_F_M≔ True "
    global switch_spat_F_M=  True
    $ 2346 "switch_spat_F_S≔ True "
    global switch_spat_F_S=  True
    $ 2347 "correction_reset()"
    correction_reset()
  elif (38 == switch_1):
    $ 2543 "Case 38"
    $ 2544 "Decap Powder container"
    $ 2545 "MoveJ"
    $ 2547 "Waypoint_7" "breakAfter"
    movej(get_inverse_kin(Waypoint_7_p, qnear=Waypoint_7_q), a=1.3962634015954636, v=1.0471975511965976, r=0.05)
    $ 2548 "MoveL"
    $ 2550 "Waypoint_8" "breakAfter"
    movel(Waypoint_8_p, a=1.2, v=0.25)
    $ 2551 "MoveL"
    $ 2552 "Decapp_above_3" "breakAfter"
    movel(Decapp_above_3_p, a=1.2, v=0.25)
    $ 2553 "Set GRP_3F_Open=On"
    set_standard_digital_out(5, True)
    $ 2554 "Wait: 0.5"
    sleep(0.5)
    $ 2555 "Decapp_place_3" "breakAfter"
    movel(Decapp_place_3_p, a=0.3, v=0.05)
    $ 2556 "Set GRP_3F_Open=Off"
    set_standard_digital_out(5, False)
    $ 2557 "Wait: 0.5"
    sleep(0.5)
    # begin: URCap Program Node
    #   Source: Robotiq_Grippers, 3.17.0.105337, Robotiq Inc.
    #   Type: Gripper
    $ 2558 "Gripper Open (1)"
    if not(gripper_connected[0]):
      popup("Gripper 1 must be connected to run this program.", "No connection", False, True, True)
    end
    if not(rq_is_gripper_activated("1")):
      popup("Gripper 1 is not activated. Go to Installation tab > Gripper to activate it and run the program again.", "Not activated", False, True, True)
    end
    rq_set_pos_spd_for(0, 77, 77, "1")
    rq_wait_pos_spe_for_request(0, 77, 77, "1")
    rq_go_to("1")
    rq_wait("1")
    # end: URCap Program Node
    $ 2559 "MoveL"
    $ 2560 "Decapp_above_4" "breakAfter"
    movel(Decapp_above_4_p, a=1.2, v=0.25)
    $ 2561 "Waypoint_78" "breakAfter"
    movel(Waypoint_78_p, a=1.2, v=0.25, r=0.05)
    $ 2562 "Home (Safe)"
    movej([-1.2302089344500047, -1.2969853503591224, -1.875639182904262, -1.539621866126728, 1.5731943360401213, -2.80099559440227], a=1.3962634015954636, v=1.0471975511965976)
  elif (39 == switch_1):
    $ 2563 "Case 39"
    $ 2564 "Powder container Pick"
    $ 2565 "Direct Pick"
    $ 2566 "Set"
    set_tcp(p[0.0,0.0,0.15052000000000001,3.1415,0.0,0.0])
    $ 2567 "read_db_data()"
    read_db_data()
    # begin: URCap Program Node
    #   Source: SensoPart VISOR Robotic, 2.0.6, SensoPart Industriesensorik GmbH
    #   Type: VISOR ChangeJob
    $ 2568 "# 1 VISOR ChangeJob"
    visor_changeJob(1, "Aztec_no_dot_pick", 6000)
    # end: URCap Program Node
    # begin: URCap Program Node
    #   Source: SensoPart VISOR Robotic, 2.0.6, SensoPart Industriesensorik GmbH
    #   Type: VISOR Terminal
    $ 2569 "# 1 VISOR Terminal"
    visor_terminal(1, "TRX00", 3000)
    # end: URCap Program Node
    $ 2570 "table_pick_TCP≔visor_getPose3d(1, 0)"
    global table_pick_TCP= visor_getPose3d (1, 0)
    # begin: URCap Program Node
    #   Source: Robotiq_Grippers, 3.17.0.105337, Robotiq Inc.
    #   Type: Gripper
    $ 2571 "Gripper Open (1)"
    if not(gripper_connected[0]):
      popup("Gripper 1 must be connected to run this program.", "No connection", False, True, True)
    end
    if not(rq_is_gripper_activated("1")):
      popup("Gripper 1 is not activated. Go to Installation tab > Gripper to activate it and run the program again.", "Not activated", False, True, True)
    end
    rq_set_pos_spd_for(0, 77, 77, "1")
    rq_wait_pos_spe_for_request(0, 77, 77, "1")
    rq_go_to("1")
    rq_wait("1")
    # end: URCap Program Node
    $ 2572 "MoveJ"
    $ 2574 "Waypoint_10" "breakAfter"
    movej(get_inverse_kin(Waypoint_10_p, qnear=Waypoint_10_q), a=1.3962634015954636, v=1.0471975511965976, r=0.05)
    $ 2575 "Waypoint_9" "breakAfter"
    movej(get_inverse_kin(Waypoint_9_p, qnear=Waypoint_9_q), a=1.3962634015954636, v=1.0471975511965976, r=0.05)
    $ 2576 "MoveJ"
    $ 2578 "table_prepick≔pose_trans(table_pick_TCP,p[0,0,cent_edge/2,0,0,0])"
    global table_prepick=pose_trans(table_pick_TCP,p[0,0,cent_edge/2,0,0,0])
    $ 2579 "table_prepick" "breakAfter"
    movej(table_prepick, a=0.8726646259971648, v=0.6981317007977318)
    $ 2580 "table_safe_pick≔pose_trans(table_prepick, p[0,pick_2_base-H_c,cent_edge/2,0,0,0])"
    global table_safe_pick= pose_trans (table_prepick, p[0,pick_2_base-H_c,cent_edge/2,0,0,0])
    $ 2581 "table_safe_pick" "breakAfter"
    movej(table_safe_pick, a=0.8726646259971648, v=0.6981317007977318, r=0.05)
    $ 2582 "table_pick≔pose_trans(table_prepick, p[0,pick_2_base - d_cc,0,0,0,0])"
    global table_pick= pose_trans (table_prepick, p[0,pick_2_base - d_cc,0,0,0,0])
    $ 2583 "table_pick" "breakAfter"
    movej(table_pick, a=0.8726646259971648, v=0.6981317007977318)
    # begin: URCap Program Node
    #   Source: Robotiq_Grippers, 3.17.0.105337, Robotiq Inc.
    #   Type: Gripper
    $ 2584 "Gripper Close (1)"
    if not(gripper_connected[0]):
      popup("Gripper 1 must be connected to run this program.", "No connection", False, True, True)
    end
    if not(rq_is_gripper_activated("1")):
      popup("Gripper 1 is not activated. Go to Installation tab > Gripper to activate it and run the program again.", "Not activated", False, True, True)
    end
    rq_set_pos_spd_for(255, 77, 51, "1")
    rq_wait_pos_spe_for_request(255, 77, 51, "1")
    rq_go_to("1")
    rq_wait("1")
    # end: URCap Program Node
    $ 2585 "table_prepick" "breakAfter"
    movej(table_prepick, a=0.8726646259971648, v=0.6981317007977318)
    $ 2586 "Picking≔ True "
    global Picking=  True
    $ 2616 "powder_position≔'Position2'"
    global powder_position="Position2"
    $ 2617 "MoveJ"
    $ 2618 "Powder_wayp1" "breakAfter"
    movej(get_inverse_kin(Powder_wayp1_p, qnear=Powder_wayp1_q), a=1.3962634015954636, v=1.0471975511965976, r=0.05)
    $ 2619 "MoveL"
    $ 2620 "Waypoint_2" "breakAfter"
    movel(Waypoint_2_p, a=1.2, v=0.25)
    $ 2621 "Set"
    set_tcp(p[0.0,0.0,0.161,3.1415,0.0,0.0])
    $ 2622 "If powder_position ≟ 'Position1'"
    if (powder_position  ==  "Position1"):
      $ 2623 "MoveJ"
      $ 2624 "Postions_otw" "breakAfter"
      movej(get_inverse_kin(Postions_otw_p, qnear=Postions_otw_q), a=1.3962634015954636, v=1.0471975511965976, r=0.01)
      $ 2625 "MoveL"
      $ 2626 "Cont_A_TCP" "breakAfter"
      movel(Cont_A_TCP, a=0.5, v=0.2)
      $ 2627 "cont_A_prepick≔pose_trans(Cont_A_TCP, p[0,0,cent_edge/2,0,0,0])"
      global cont_A_prepick= pose_trans (Cont_A_TCP, p[0,0,cent_edge/2,0,0,0])
      $ 2628 "cont_A_prepick" "breakAfter"
      movel(cont_A_prepick, a=0.3, v=0.05)
      $ 2629 "cont_A_pick≔pose_trans(cont_A_prepick, p[0,pick_2_base-d_cc,0,0,0,0])"
      global cont_A_pick= pose_trans (cont_A_prepick, p[0,pick_2_base-d_cc,0,0,0,0])
      $ 2630 "cont_A_pick" "breakAfter"
      movel(cont_A_pick, a=0.2, v=0.1)
      # begin: URCap Program Node
      #   Source: Robotiq_Grippers, 3.17.0.105337, Robotiq Inc.
      #   Type: Gripper
      $ 2631 "Gripper Open (1)"
      if not(gripper_connected[0]):
        popup("Gripper 1 must be connected to run this program.", "No connection", False, True, True)
      end
      if not(rq_is_gripper_activated("1")):
        popup("Gripper 1 is not activated. Go to Installation tab > Gripper to activate it and run the program again.", "Not activated", False, True, True)
      end
      rq_set_pos_spd_for(0, 77, 26, "1")
      rq_wait_pos_spe_for_request(0, 77, 26, "1")
      rq_go_to("1")
      rq_wait("1")
      # end: URCap Program Node
      $ 2632 "cont_A_otw" "breakAfter"
      movel(cont_A_otw_p, a=0.5, v=0.2)
      $ 2633 "cont_A_prepick" "breakAfter"
      movel(cont_A_prepick, a=0.5, v=0.2)
      $ 2634 "Postions_otw" "breakAfter"
      movel(Postions_otw_p, a=0.5, v=0.2, r=0.01)
      $ 2636 "Home (Safe)"
      movej([-1.2302089344500047, -1.2969853503591224, -1.875639182904262, -1.539621866126728, 1.5731943360401213, -2.80099559440227], a=1.3962634015954636, v=1.0471975511965976)
    else:
      $ 2638 "ElseIf powder_position≟'Position2'"
      if (powder_position == "Position2"):
        $ 2639 "MoveJ"
        $ 2640 "Postions_otw" "breakAfter"
        movej(get_inverse_kin(Postions_otw_p, qnear=Postions_otw_q), a=1.3962634015954636, v=1.0471975511965976, r=0.01)
        $ 2641 "MoveL"
        $ 2644 "cont_B_prepick≔pose_trans(Cont_B_TCP, p[0,0,cent_edge/2,0,0,0])"
        global cont_B_prepick= pose_trans (Cont_B_TCP, p[0,0,cent_edge/2,0,0,0])
        $ 2645 "cont_B_prepick" "breakAfter"
        movel(cont_B_prepick, a=1.2, v=0.25)
        $ 2646 "cont_B_pick≔pose_trans(cont_B_prepick, p[0,pick_2_base-d_cc,0,0,0,0])"
        global cont_B_pick= pose_trans (cont_B_prepick, p[0,pick_2_base-d_cc,0,0,0,0])
        $ 2647 "cont_B_pick" "breakAfter"
        global move_thread_flag_2647=0
        thread move_thread_2647():
          enter_critical
          move_thread_flag_2647 = 1
          movel(cont_B_pick, a=0.2, v=0.1)
          move_thread_flag_2647 = 2
          exit_critical
        end
        move_thread_flag_2647 = 0
        move_thread_han_2647 = run move_thread_2647()
        while (True):
          local targetTcpDirection=get_target_tcp_speed()
          local stepsToRetract=tool_contact(direction=targetTcpDirection, force_threshold=8.000000)
          if (stepsToRetract > 0):
            kill move_thread_han_2647
            stopl(3.0)
            local backTrackMovement=get_actual_joint_positions_history(stepsToRetract)
            local contactPose=get_forward_kin(backTrackMovement)
            local posDir=[targetTcpDirection[0],targetTcpDirection[1],targetTcpDirection[2]]
            local retractTo=contactPose
            if (norm(posDir) > 1e-6):
              local normalizedPosDir=normalize(posDir)
              local additionalRetraction=p[normalizedPosDir[0] * 0.0, normalizedPosDir[1] * 0.0, normalizedPosDir[2] * 0.0, 0, 0, 0]
              retractTo = pose_sub(contactPose, additionalRetraction)
            end
            movel(retractTo, a=3.0, v=0.1)
            $ 2648 "Until (tool_contact_detection)"
            $ 2649 "saved_place_pos≔get_actual_tcp_pose()"
            global saved_place_pos= get_actual_tcp_pose ()
            break
          end
          sleep(1.0E-10)
          if (move_thread_flag_2647 > 1):
            join move_thread_han_2647
            break
          end
          sync()
        end
        # begin: URCap Program Node
        #   Source: Robotiq_Grippers, 3.17.0.105337, Robotiq Inc.
        #   Type: Gripper
        $ 2650 "Gripper Open (1)"
        if not(gripper_connected[0]):
          popup("Gripper 1 must be connected to run this program.", "No connection", False, True, True)
        end
        if not(rq_is_gripper_activated("1")):
          popup("Gripper 1 is not activated. Go to Installation tab > Gripper to activate it and run the program again.", "Not activated", False, True, True)
        end
        rq_set_pos_spd_for(0, 77, 26, "1")
        rq_wait_pos_spe_for_request(0, 77, 26, "1")
        rq_go_to("1")
        rq_wait("1")
        # end: URCap Program Node
        $ 2651 "cont_B_otw" "breakAfter"
        movel(cont_B_otw_p, a=1.2, v=0.25)
        $ 2653 "cont_B_safe" "breakAfter"
        movel(cont_B_safe_p, a=1.2, v=0.25)
        $ 2654 "Postions_otw" "breakAfter"
        movel(Postions_otw_p, a=1.2, v=0.25)
        $ 2655 "Home (Safe)"
        movej([-1.2302089344500047, -1.2969853503591224, -1.875639182904262, -1.539621866126728, 1.5731943360401213, -2.80099559440227], a=1.3962634015954636, v=1.0471975511965976)
      else:
        $ 2657 "ElseIf powder_position≟'Position3'"
        if (powder_position == "Position3"):
          $ 2658 "MoveJ"
          $ 2659 "Postions_otw" "breakAfter"
          movej(get_inverse_kin(Postions_otw_p, qnear=Postions_otw_q), a=1.3962634015954636, v=1.0471975511965976, r=0.01)
          $ 2666 "MoveL"
          $ 2667 "Cont_C_TCP" "breakAfter"
          movel(Cont_C_TCP, a=1.2, v=0.25, r=0.01)
          $ 2668 "cont_C_prepick≔pose_trans(Cont_C_TCP, p[0,0,cent_edge/2,0,0,0])"
          global cont_C_prepick= pose_trans (Cont_C_TCP, p[0,0,cent_edge/2,0,0,0])
          $ 2669 "cont_C_prepick" "breakAfter"
          movel(cont_C_prepick, a=0.3, v=0.05)
          $ 2670 "cont_C_pick≔pose_trans(cont_C_prepick, p[0,pick_2_base-d_cc,0,0,0,0])"
          global cont_C_pick= pose_trans (cont_C_prepick, p[0,pick_2_base-d_cc,0,0,0,0])
          $ 2671 "cont_C_pick" "breakAfter"
          movel(cont_C_pick, a=0.2, v=0.1)
          # begin: URCap Program Node
          #   Source: Robotiq_Grippers, 3.17.0.105337, Robotiq Inc.
          #   Type: Gripper
          $ 2672 "Gripper Open (1)"
          if not(gripper_connected[0]):
            popup("Gripper 1 must be connected to run this program.", "No connection", False, True, True)
          end
          if not(rq_is_gripper_activated("1")):
            popup("Gripper 1 is not activated. Go to Installation tab > Gripper to activate it and run the program again.", "Not activated", False, True, True)
          end
          rq_set_pos_spd_for(0, 77, 26, "1")
          rq_wait_pos_spe_for_request(0, 77, 26, "1")
          rq_go_to("1")
          rq_wait("1")
          # end: URCap Program Node
          $ 2673 "cont_C_otw" "breakAfter"
          movel(cont_C_otw_p, a=1.2, v=0.25)
          $ 2674 "cont_C_prepick" "breakAfter"
          movel(cont_C_prepick, a=1.2, v=0.25, r=0.01)
          $ 2675 "Postions_otw" "breakAfter"
          movel(Postions_otw_p, a=1.2, v=0.25)
          $ 2676 "Home (Safe)"
          movej([-1.2302089344500047, -1.2969853503591224, -1.875639182904262, -1.539621866126728, 1.5731943360401213, -2.80099559440227], a=1.3962634015954636, v=1.0471975511965976)
        end
      end
    end
    $ 2678 "Home (Safe)"
    movej([-1.2302089344500047, -1.2969853503591224, -1.875639182904262, -1.539621866126728, 1.5731943360401213, -2.80099559440227], a=1.3962634015954636, v=1.0471975511965976)
  elif (41 == switch_1):
    $ 2787 "Case 41"
    $ 2788 "Task≔'Decapping_Dosing'"
    global Task="Decapping_Dosing"
    $ 2789 "tilt_to_home()"
    tilt_to_home()
    $ 2790 "Weigh, Place & decap container"
    $ 2791 "Set"
    set_tcp(p[0.0,0.0,0.15052000000000001,3.1415,0.0,0.0])
    # begin: URCap Program Node
    #   Source: SensoPart VISOR Robotic, 2.0.6, SensoPart Industriesensorik GmbH
    #   Type: VISOR Robotic App
    $ 2792 "VISOR Easy Pick"
    def visorFuncEasyPick_66369a():
      # begin: URCap Program Node
      #   Source: SensoPart VISOR Robotic, 2.0.6, SensoPart Industriesensorik GmbH
      #   Type: Easy Pick Setup
      $ 2793 "# 1 Setup" "noBreak"
      local easyPickVisorId = 1
      local easyPickArmMounted = True
      local easyPickSetJob = True
      local easyPickJobName = "PoTS"
      local easyPickAtImgAcq = False
      local easyPickImgAcqPose = FRM_PoTS
      # end: URCap Program Node
      # begin: URCap Program Node
      #   Source: SensoPart VISOR Robotic, 2.0.6, SensoPart Industriesensorik GmbH
      #   Type: Process
      $ 2794 "Process" "noBreak"
      local easyPickObjTaken = False
      local easyPickTrigger = False
      local easyPickPoseIdx = 0
      local easyPickPose = p[0,0,0,0,0,0]
      def easyPickFuncTrigger(visorId, setJob, jobName, arm):
      if (setJob):
        visor_changeJob(visorId, jobName, 6000)
      end
      if (arm):
        visor_trigger(visorId, 6000, "arm")
      else:
        visor_trigger(visorId, 6000)
      end
      global easyPickParts_7=visor_partsFound(visorId)
      visor_easyPickUpdate(visorId, "parts", visor_partsFound(visorId))
      return visor_getPose3d(visorId, 0)
    end
    while (not easyPickObjTaken):
      easyPickTrigger = (easyPickCount_7 >= visor_partsFound(easyPickVisorId)) or (easyPickCount_7 > 9) or (not visor_easyPickCheckIdent("b73a64", easyPickVisorId))
      if (easyPickTrigger):
        easyPickCount_7 = 0
      end
      easyPickPoseIdx = easyPickCount_7
      easyPickPose = visor_getPose3d(easyPickVisorId, easyPickPoseIdx)
      visor_easyPickUpdate(easyPickVisorId, "counter", easyPickPoseIdx)
      # begin: URCap Program Node
      #   Source: SensoPart VISOR Robotic, 2.0.6, SensoPart Industriesensorik GmbH
      #   Type: Image Acquisition Pose
      $ 2795 "Image Acquisition Pose" "noBreak"
      if (easyPickTrigger):
        if (not easyPickAtImgAcq):
          movej(pose_trans(easyPickImgAcqPose,p[0.0000,0.0000,-0.0000,0.0000,0.0000,0.0000]),a=1.3963,v=1.0472,t=0.000000,r=0.000000)
          easyPickAtImgAcq = True
        end
        easyPickPose = easyPickFuncTrigger(easyPickVisorId, easyPickSetJob, easyPickJobName, easyPickArmMounted)
      end
      # end: URCap Program Node
      # begin: URCap Program Node
      #   Source: SensoPart VISOR Robotic, 2.0.6, SensoPart Industriesensorik GmbH
      #   Type: Object Detected
      $ 2796 "Object Detected" "noBreak"
      if (visor_partsFound(easyPickVisorId) > 0):
        $ 2797 "Open Gripper" "noBreak"
        # begin: URCap Program Node
        #   Source: Robotiq_Grippers, 3.17.0.105337, Robotiq Inc.
        #   Type: Gripper
        $ 2798 "Gripper Open (1)" "noBreak"
        if not(gripper_connected[0]):
          popup("Gripper 1 must be connected to run this program.", "No connection", False, True, True)
        end
        if not(rq_is_gripper_activated("1")):
          popup("Gripper 1 is not activated. Go to Installation tab > Gripper to activate it and run the program again.", "Not activated", False, True, True)
        end
        rq_set_pos_spd_for(0, 77, 77, "1")
        rq_wait_pos_spe_for_request(0, 77, 77, "1")
        rq_go_to("1")
        rq_wait("1")
        # end: URCap Program Node
        $ 2799 "Set" "noBreak"
        set_tcp(p[0.0,0.0,0.161,3.1415,0.0,0.0])
        $ 2800 "Wait: 0.2" "noBreak"
        sleep(0.2)
        $ 2801 "Place on second weigh scale" "noBreak"
        $ 2802 "MoveJ" "noBreak"
        $ 2803 "Waypoint_1" "noBreak"
        movej(get_inverse_kin(Waypoint_1_p, qnear=Waypoint_1_q), a=1.3962634015954636, v=1.0471975511965976, r=0.1)
        $ 2804 "Waypoint_5" "noBreak"
        movej(get_inverse_kin(Waypoint_5_p, qnear=Waypoint_5_q), a=1.3962634015954636, v=1.0471975511965976)
        $ 2806 "If Picking≟ True " "noBreak"
        if (Picking ==   True  ):
          $ 2807 "Pick from saved pose" "noBreak"
          $ 2808 "MoveL" "noBreak"
          $ 2809 "cont_B_safe" "noBreak"
          movel(cont_B_safe_p, a=0.2, v=0.1)
          $ 2810 "saved_place_pos" "noBreak"
          movel(saved_place_pos, a=1.2, v=0.25)
          # begin: URCap Program Node
          #   Source: Robotiq_Grippers, 3.17.0.105337, Robotiq Inc.
          #   Type: Gripper
          $ 2811 "Gripper Close (1)" "noBreak"
          if not(gripper_connected[0]):
            popup("Gripper 1 must be connected to run this program.", "No connection", False, True, True)
          end
          if not(rq_is_gripper_activated("1")):
            popup("Gripper 1 is not activated. Go to Installation tab > Gripper to activate it and run the program again.", "Not activated", False, True, True)
          end
          rq_set_pos_spd_for(255, 77, 26, "1")
          rq_wait_pos_spe_for_request(255, 77, 26, "1")
          rq_go_to("1")
          rq_wait("1")
          # end: URCap Program Node
          $ 2812 "cont_B_safe" "noBreak"
          movel(cont_B_safe_p, a=1.2, v=0.25)
          $ 2813 "Postions_otw" "noBreak"
          movel(Postions_otw_p, a=1.2, v=0.25)
        else:
          $ 2816 "Else" "noBreak"
          $ 2817 "read_db_data()" "noBreak"
          read_db_data()
          $ 2818 "Pick from B" "noBreak"
          $ 2819 "MoveL" "noBreak"
          $ 2821 "cont_B_safe" "noBreak"
          movel(cont_B_safe_p, a=1.2, v=0.25)
          $ 2822 "cont_B_prepick≔pose_trans(Cont_B_TCP, p[0,0,cent_edge/2,0,0,0])" "noBreak"
          global cont_B_prepick= pose_trans (Cont_B_TCP, p[0,0,cent_edge/2,0,0,0])
          $ 2823 "cont_B_otw" "noBreak"
          movel(cont_B_otw_p, a=1.2, v=0.25)
          $ 2825 "cont_B_pick≔pose_trans(cont_B_prepick, p[0,pick_2_base-d_cc,0,0,0,0])" "noBreak"
          global cont_B_pick= pose_trans (cont_B_prepick, p[0,pick_2_base-d_cc,0,0,0,0])
          $ 2826 "cont_B_pick" "noBreak"
          movel(cont_B_pick, a=0.2, v=0.1)
          # begin: URCap Program Node
          #   Source: Robotiq_Grippers, 3.17.0.105337, Robotiq Inc.
          #   Type: Gripper
          $ 2827 "Gripper Close (1)" "noBreak"
          if not(gripper_connected[0]):
            popup("Gripper 1 must be connected to run this program.", "No connection", False, True, True)
          end
          if not(rq_is_gripper_activated("1")):
            popup("Gripper 1 is not activated. Go to Installation tab > Gripper to activate it and run the program again.", "Not activated", False, True, True)
          end
          rq_set_pos_spd_for(255, 77, 51, "1")
          rq_wait_pos_spe_for_request(255, 77, 51, "1")
          rq_go_to("1")
          rq_wait("1")
          # end: URCap Program Node
          $ 2828 "cont_B_prepick" "noBreak"
          movel(cont_B_prepick, a=1.2, v=0.25, r=0.01)
          $ 2829 "Postions_otw" "noBreak"
          movel(Postions_otw_p, a=1.2, v=0.25)
        end
        $ 2846 "Set" "noBreak"
        set_tcp(p[0.0,0.0,0.15052000000000001,3.1415,0.0,0.0])
        # begin: URCap Program Node
        #   Source: SensoPart VISOR Robotic, 2.0.6, SensoPart Industriesensorik GmbH
        #   Type: Approach Pose
        $ 2847 "Approach Pose" "noBreak"
        movej(pose_trans(easyPickPose,p[0.0000,0.0000,-0.0000,0.0000,0.0000,0.0000]),a=0.5236,v=0.4363,t=0.000000,r=0.000000)
        # end: URCap Program Node
        # begin: URCap Program Node
        #   Source: SensoPart VISOR Robotic, 2.0.6, SensoPart Industriesensorik GmbH
        #   Type: Target Pose
        $ 2848 "Target Pose" "noBreak"
        movel(pose_trans(easyPickPose,p[0.0000,0.0000,-0.0000,0.0000,0.0000,0.0000]),a=0.1000,v=0.0500,t=0.000000,r=0.000000)
        # end: URCap Program Node
        $ 2849 "Close Gripper" "noBreak"
        $ 2850 "container_place≔get_actual_tcp_pose()" "noBreak"
        global container_place= get_actual_tcp_pose ()
        $ 2851 "PoTS_place_abov≔pose_trans(container_place, p[0,0,cent_edge/2,0,0,0])" "noBreak"
        global PoTS_place_abov=pose_trans(container_place, p[0,0,cent_edge/2,0,0,0])
        $ 2852 "MoveL" "noBreak"
        $ 2853 "PoTS_place_abov" "noBreak"
        movel(PoTS_place_abov, a=0.5, v=0.05)
        $ 2855 "target_pose≔pose_trans(PoTS_place_abov, p[0,pick_2_base-d_cc,0,0,0,0])" "noBreak"
        global target_pose=pose_trans(PoTS_place_abov, p[0,pick_2_base-d_cc,0,0,0,0])
        $ 2856 "MoveL" "noBreak"
        $ 2857 "target_pose" "noBreak"
        movel(target_pose, a=0.3, v=0.05)
        # begin: URCap Program Node
        #   Source: Robotiq_Grippers, 3.17.0.105337, Robotiq Inc.
        #   Type: Gripper
        $ 2858 "Gripper Open (1)" "noBreak"
        if not(gripper_connected[0]):
          popup("Gripper 1 must be connected to run this program.", "No connection", False, True, True)
        end
        if not(rq_is_gripper_activated("1")):
          popup("Gripper 1 is not activated. Go to Installation tab > Gripper to activate it and run the program again.", "Not activated", False, True, True)
        end
        rq_set_pos_spd_for(0, 77, 77, "1")
        rq_wait_pos_spe_for_request(0, 77, 77, "1")
        rq_go_to("1")
        rq_wait("1")
        # end: URCap Program Node
        # begin: URCap Program Node
        #   Source: SensoPart VISOR Robotic, 2.0.6, SensoPart Industriesensorik GmbH
        #   Type: Exit Pose
        $ 2859 "Exit Pose" "noBreak"
        movel(pose_trans(easyPickPose,p[0.0000,0.0000,0.1000,0.0000,0.0000,0.0000]),a=0.5000,v=0.2500,t=0.000000,r=0.000000)
        # end: URCap Program Node
        easyPickObjTaken = True
      end
      # end: URCap Program Node
      # begin: URCap Program Node
      #   Source: SensoPart VISOR Robotic, 2.0.6, SensoPart Industriesensorik GmbH
      #   Type: No Object Detected
      $ 2860 "No Object Detected" "noBreak"
      if (visor_partsFound(easyPickVisorId) < 1):
        $ 2861 "Popup: No POTS detected" "noBreak"
        popup("No POTS detected", "Message", False, False, blocking=True)
        else:
      end
      # end: URCap Program Node
    end
    easyPickCount_7 = easyPickCount_7 + 1
    visor_easyPickUpdate(easyPickVisorId, "counter", easyPickCount_7)
    visor_easyPickSetIdent("b73a64", easyPickVisorId)
    # end: URCap Program Node
  end
  visorFuncEasyPick_66369a()
  # end: URCap Program Node
  $ 2896 "MoveJ"
  $ 2897 "place_2_home" "breakAfter"
  movej(get_inverse_kin(place_2_home_p, qnear=place_2_home_q), a=1.3962634015954636, v=1.0471975511965976)
  $ 2898 "Picking≔ False "
  global Picking=  False
  elif (42 == switch_1):
    $ 2899 "Case 42"
  elif (43 == switch_1):
    $ 3661 "Case 43"
  elif (44 == switch_1):
    $ 3914 "Case 44"
  elif (45 == switch_1):
    $ 3978 "Case 45"
  elif (46 == switch_1):
    $ 4015 "Case 46"
  elif (47 == switch_1):
    $ 4305 "Case 47"
  elif (48 == switch_1):
    $ 4360 "Case 48"
  elif (49 == switch_1):
    $ 4378 "Case 49"
  elif (50 == switch_1):
    $ 4396 "Case 50"
    $ 4397 "Emptying powder container"
    $ 4398 "tilt_to_home()"
    tilt_to_home()
    $ 4399 "scoop_status≔'emptying'"
    global scoop_status="emptying"
    $ 4400 "Dosing untill empty"
    $ 4401 "tilt_angle_sent≔0.0"
    global tilt_angle_sent=0.0
    $ 4402 "send_target_info()"
    send_target_info()
    $ 4403 "zero_scale()"
    zero_scale()
    $ 4404 "prev_spat≔''"
    global prev_spat=""
    $ 4405 "spatula≔''"
    global spatula=""
    $ 4406 "send_powder_info()"
    send_powder_info()
    $ 4407 "Set AO[0]=0.0"
    set_standard_analog_out(0, 0.0)
    $ 4408 "Wait: 0.2"
    sleep(0.2)
    $ 4409 "reach pots decapping pose"
    # begin: URCap Program Node
    #   Source: SensoPart VISOR Robotic, 2.0.6, SensoPart Industriesensorik GmbH
    #   Type: VISOR Robotic App
    $ 4415 "VISOR Easy Pick"
    def visorFuncEasyPick_b3e024():
      # begin: URCap Program Node
      #   Source: SensoPart VISOR Robotic, 2.0.6, SensoPart Industriesensorik GmbH
      #   Type: Easy Pick Setup
      $ 4416 "# 1 Setup" "noBreak"
      local easyPickVisorId = 1
      local easyPickArmMounted = True
      local easyPickSetJob = True
      local easyPickJobName = "Weight_scale"
      local easyPickAtImgAcq = False
      local easyPickImgAcqPose = Trigger
      # end: URCap Program Node
      # begin: URCap Program Node
      #   Source: SensoPart VISOR Robotic, 2.0.6, SensoPart Industriesensorik GmbH
      #   Type: Process
      $ 4417 "Process" "noBreak"
      local easyPickObjTaken = False
      local easyPickTrigger = False
      local easyPickPoseIdx = 0
      local easyPickPose = p[0,0,0,0,0,0]
      def easyPickFuncTrigger(visorId, setJob, jobName, arm):
      if (setJob):
        visor_changeJob(visorId, jobName, 6000)
      end
      if (arm):
        visor_trigger(visorId, 6000, "arm")
      else:
        visor_trigger(visorId, 6000)
      end
      global easyPickParts_4=visor_partsFound(visorId)
      visor_easyPickUpdate(visorId, "parts", visor_partsFound(visorId))
      return visor_getPose3d(visorId, 0)
    end
    while (not easyPickObjTaken):
      easyPickTrigger = (easyPickCount_4 >= visor_partsFound(easyPickVisorId)) or (easyPickCount_4 > 9) or (not visor_easyPickCheckIdent("cf8854", easyPickVisorId))
      if (easyPickTrigger):
        easyPickCount_4 = 0
      end
      easyPickPoseIdx = easyPickCount_4
      easyPickPose = visor_getPose3d(easyPickVisorId, easyPickPoseIdx)
      visor_easyPickUpdate(easyPickVisorId, "counter", easyPickPoseIdx)
      # begin: URCap Program Node
      #   Source: SensoPart VISOR Robotic, 2.0.6, SensoPart Industriesensorik GmbH
      #   Type: Image Acquisition Pose
      $ 4418 "Image Acquisition Pose" "noBreak"
      if (easyPickTrigger):
        if (not easyPickAtImgAcq):
          movej(pose_trans(easyPickImgAcqPose,p[0.0000,0.0000,-0.0000,0.0000,0.0000,0.0000]),a=1.3963,v=1.0472,t=0.000000,r=0.000000)
          easyPickAtImgAcq = True
        end
        easyPickPose = easyPickFuncTrigger(easyPickVisorId, easyPickSetJob, easyPickJobName, easyPickArmMounted)
      end
      # end: URCap Program Node
      # begin: URCap Program Node
      #   Source: SensoPart VISOR Robotic, 2.0.6, SensoPart Industriesensorik GmbH
      #   Type: Object Detected
      $ 4419 "Object Detected" "noBreak"
      if (visor_partsFound(easyPickVisorId) > 0):
        $ 4420 "Open Gripper" "noBreak"
        $ 4421 "weight_value≔get_weight()" "noBreak"
        global weight_value=get_weight()
        $ 4422 "Wait: 1.0" "noBreak"
        sleep(1.0)
        $ 4423 "diff≔target_weight-weight_value" "noBreak"
        global diff=target_weight-weight_value
        $ 4424 "compute_level_percent(W_now, weight_value)" "noBreak"
        compute_level_percent(W_now, weight_value)
        $ 4425 "send_level_info()" "noBreak"
        send_level_info()
        $ 4426 "spatula≔select_spatula(Flowability, level, diff, bulk_density, mouth_d)" "noBreak"
        global spatula=select_spatula(Flowability, level, diff, bulk_density, mouth_d)
        $ 4427 "Wait: 0.2" "noBreak"
        sleep(0.2)
        $ 4428 "send_spatula_info()" "noBreak"
        send_spatula_info()
        $ 4429 "Pick spatula" "noBreak"
        $ 4430 "If spatula ≟ 'spatula_L'" "noBreak"
        if (spatula  ==  "spatula_L"):
          $ 4431 "MoveJ" "noBreak"
          $ 4432 "Spatula_otw" "noBreak"
          movej(get_inverse_kin(Spatula_otw_p, qnear=Spatula_otw_q), a=1.3962634015954636, v=1.0471975511965976)
          $ 4433 "pick_spat_L_abv" "noBreak"
          movej(get_inverse_kin(pick_spat_L_abv_p, qnear=pick_spat_L_abv_q), a=1.3962634015954636, v=1.0471975511965976)
          $ 4434 "MoveL" "noBreak"
          $ 4435 "spat_L_pick" "noBreak"
          movel(spat_L_pick_p, a=1.2, v=0.25)
          # begin: URCap Program Node
          #   Source: Robotiq_Grippers, 3.17.0.105337, Robotiq Inc.
          #   Type: Gripper
          $ 4436 "Gripper Close (1)" "noBreak"
          if not(gripper_connected[0]):
            popup("Gripper 1 must be connected to run this program.", "No connection", False, True, True)
          end
          if not(rq_is_gripper_activated("1")):
            popup("Gripper 1 is not activated. Go to Installation tab > Gripper to activate it and run the program again.", "Not activated", False, True, True)
          end
          rq_set_pos_spd_for(255, 0, 77, "1")
          rq_wait_pos_spe_for_request(255, 0, 77, "1")
          rq_go_to("1")
          rq_wait("1")
          # end: URCap Program Node
          $ 4437 "spat_L_lift" "noBreak"
          movel(spat_L_lift_p, a=1.2, v=0.25, r=0.01)
          $ 4438 "spat_L_side" "noBreak"
          movel(spat_L_side_p, a=1.2, v=0.25, r=0.01)
          $ 4439 "spat_L_up" "noBreak"
          movel(spat_L_up_p, a=1.2, v=0.25, r=0.05)
          $ 4440 "MoveJ" "noBreak"
          $ 4441 "Spatula_otw" "noBreak"
          movej(get_inverse_kin(Spatula_otw_p, qnear=Spatula_otw_q), a=1.3962634015954636, v=1.0471975511965976)
        else:
          $ 4442 "ElseIf spatula ≟'spatula_M'" "noBreak"
          if (spatula  == "spatula_M"):
            $ 4443 "MoveJ" "noBreak"
            $ 4444 "Spatula_otw" "noBreak"
            movej(get_inverse_kin(Spatula_otw_p, qnear=Spatula_otw_q), a=1.3962634015954636, v=1.0471975511965976)
            $ 4445 "spat_M_up" "noBreak"
            movej(get_inverse_kin(spat_M_up_p, qnear=spat_M_up_q), a=1.3962634015954636, v=1.0471975511965976, r=0.05)
            $ 4446 "MoveL" "noBreak"
            $ 4447 "spat_M_pick" "noBreak"
            movel(spat_M_pick_p, a=1.2, v=0.25)
            # begin: URCap Program Node
            #   Source: Robotiq_Grippers, 3.17.0.105337, Robotiq Inc.
            #   Type: Gripper
            $ 4448 "Gripper Close (1)" "noBreak"
            if not(gripper_connected[0]):
              popup("Gripper 1 must be connected to run this program.", "No connection", False, True, True)
            end
            if not(rq_is_gripper_activated("1")):
              popup("Gripper 1 is not activated. Go to Installation tab > Gripper to activate it and run the program again.", "Not activated", False, True, True)
            end
            rq_set_pos_spd_for(255, 0, 77, "1")
            rq_wait_pos_spe_for_request(255, 0, 77, "1")
            rq_go_to("1")
            rq_wait("1")
            # end: URCap Program Node
            $ 4449 "spat_M_up" "noBreak"
            movel(spat_M_up_p, a=1.2, v=0.25, r=0.05)
            $ 4450 "Spatula_otw" "noBreak"
            movel(Spatula_otw_p, a=1.2, v=0.25)
            $ 4451 "switch_spat_M≔ False " "noBreak"
            global switch_spat_M=  False
          else:
            $ 4452 "ElseIf spatula≟'spatula_S'" "noBreak"
            if (spatula == "spatula_S"):
              $ 4453 "MoveJ" "noBreak"
              $ 4454 "Spatula_otw" "noBreak"
              movej(get_inverse_kin(Spatula_otw_p, qnear=Spatula_otw_q), a=1.3962634015954636, v=1.0471975511965976)
              $ 4455 "spat_S_Up_7" "noBreak"
              movej(get_inverse_kin(spat_S_Up_7_p, qnear=spat_S_Up_7_q), a=1.3962634015954636, v=1.0471975511965976, r=0.05)
              $ 4456 "MoveL" "noBreak"
              $ 4457 "spat_S_Pick_4" "noBreak"
              movel(spat_S_Pick_4_p, a=1.2, v=0.25)
              # begin: URCap Program Node
              #   Source: Robotiq_Grippers, 3.17.0.105337, Robotiq Inc.
              #   Type: Gripper
              $ 4458 "Gripper Close (1)" "noBreak"
              if not(gripper_connected[0]):
                popup("Gripper 1 must be connected to run this program.", "No connection", False, True, True)
              end
              if not(rq_is_gripper_activated("1")):
                popup("Gripper 1 is not activated. Go to Installation tab > Gripper to activate it and run the program again.", "Not activated", False, True, True)
              end
              rq_set_pos_spd_for(255, 0, 77, "1")
              rq_wait_pos_spe_for_request(255, 0, 77, "1")
              rq_go_to("1")
              rq_wait("1")
              # end: URCap Program Node
              $ 4459 "spat_S_Up_8" "noBreak"
              movel(spat_S_Up_8_p, a=1.2, v=0.25, r=0.05)
              $ 4460 "Spatula_otw" "noBreak"
              movel(Spatula_otw_p, a=1.2, v=0.25)
              $ 4461 "switch_spat_S≔ False " "noBreak"
              global switch_spat_S=  False
            else:
              $ 4462 "ElseIf spatula≟'spatula_flat_M'" "noBreak"
              if (spatula == "spatula_flat_M"):
                $ 4463 "MoveJ" "noBreak"
                $ 4464 "Spatula_otw" "noBreak"
                movej(get_inverse_kin(Spatula_otw_p, qnear=Spatula_otw_q), a=1.3962634015954636, v=1.0471975511965976)
                $ 4465 "spat_flatM_up" "noBreak"
                movej(get_inverse_kin(spat_flatM_up_p, qnear=spat_flatM_up_q), a=1.3962634015954636, v=1.0471975511965976, r=0.05)
                $ 4466 "MoveL" "noBreak"
                $ 4467 "spat_flatM_pick" "noBreak"
                movel(spat_flatM_pick_p, a=1.2, v=0.25)
                # begin: URCap Program Node
                #   Source: Robotiq_Grippers, 3.17.0.105337, Robotiq Inc.
                #   Type: Gripper
                $ 4468 "Gripper Close (1)" "noBreak"
                if not(gripper_connected[0]):
                  popup("Gripper 1 must be connected to run this program.", "No connection", False, True, True)
                end
                if not(rq_is_gripper_activated("1")):
                  popup("Gripper 1 is not activated. Go to Installation tab > Gripper to activate it and run the program again.", "Not activated", False, True, True)
                end
                rq_set_pos_spd_for(255, 0, 77, "1")
                rq_wait_pos_spe_for_request(255, 0, 77, "1")
                rq_go_to("1")
                rq_wait("1")
                # end: URCap Program Node
                $ 4469 "spat_flatM_up" "noBreak"
                movel(spat_flatM_up_p, a=1.2, v=0.25, r=0.05)
                $ 4470 "Spatula_otw" "noBreak"
                movel(Spatula_otw_p, a=1.2, v=0.25)
                $ 4471 "switch_spat_F_M≔ False " "noBreak"
                global switch_spat_F_M=  False
              else:
                $ 4472 "ElseIf spatula≟'spatula_flat_S'" "noBreak"
                if (spatula == "spatula_flat_S"):
                  $ 4473 "MoveJ" "noBreak"
                  $ 4474 "Spatula_otw" "noBreak"
                  movej(get_inverse_kin(Spatula_otw_p, qnear=Spatula_otw_q), a=1.3962634015954636, v=1.0471975511965976)
                  $ 4475 "spat_flatS_up" "noBreak"
                  movej(get_inverse_kin(spat_flatS_up_p, qnear=spat_flatS_up_q), a=1.3962634015954636, v=1.0471975511965976, r=0.05)
                  $ 4476 "MoveL" "noBreak"
                  $ 4477 "spat_flatS_pick" "noBreak"
                  movel(spat_flatS_pick_p, a=1.2, v=0.25)
                  # begin: URCap Program Node
                  #   Source: Robotiq_Grippers, 3.17.0.105337, Robotiq Inc.
                  #   Type: Gripper
                  $ 4478 "Gripper Close (1)" "noBreak"
                  if not(gripper_connected[0]):
                    popup("Gripper 1 must be connected to run this program.", "No connection", False, True, True)
                  end
                  if not(rq_is_gripper_activated("1")):
                    popup("Gripper 1 is not activated. Go to Installation tab > Gripper to activate it and run the program again.", "Not activated", False, True, True)
                  end
                  rq_set_pos_spd_for(255, 0, 77, "1")
                  rq_wait_pos_spe_for_request(255, 0, 77, "1")
                  rq_go_to("1")
                  rq_wait("1")
                  # end: URCap Program Node
                  $ 4479 "spat_flatS_up" "noBreak"
                  movel(spat_flatS_up_p, a=1.2, v=0.25, r=0.05)
                  $ 4480 "Spatula_otw" "noBreak"
                  movel(Spatula_otw_p, a=1.2, v=0.25)
                  $ 4481 "switch_spat_F_S≔ False " "noBreak"
                  global switch_spat_F_S=  False
                end
              end
            end
          end
        end
        $ 4482 "Action_Info≔'Scooping'" "noBreak"
        global Action_Info="Scooping"
        $ 4483 "auto_tilt_and_scoop(W_now, target_weight, weight_value)" "noBreak"
        auto_tilt_and_scoop(W_now, target_weight, weight_value)
        $ 4484 "Action_Info≔'Dosing'" "noBreak"
        global Action_Info="Dosing"
        # begin: URCap Program Node
        #   Source: SensoPart VISOR Robotic, 2.0.6, SensoPart Industriesensorik GmbH
        #   Type: Approach Pose
        $ 4485 "Approach Pose" "noBreak"
        movej(pose_trans(easyPickPose,p[0.0000,0.0000,-0.0000,0.0000,0.0000,0.0000]),a=0.2618,v=0.1745,t=0.000000,r=0.000000)
        # end: URCap Program Node
        # begin: URCap Program Node
        #   Source: SensoPart VISOR Robotic, 2.0.6, SensoPart Industriesensorik GmbH
        #   Type: Target Pose
        $ 4486 "Target Pose" "noBreak"
        movel(pose_trans(easyPickPose,p[0.0000,0.0000,-0.0000,0.0000,0.0000,0.0000]),a=0.0500,v=0.0200,t=0.000000,r=0.000000)
        # end: URCap Program Node
        $ 4487 "Close Gripper" "noBreak"
        $ 4488 "dispense_pos≔get_actual_tcp_pose()" "noBreak"
        global dispense_pos= get_actual_tcp_pose ()
        $ 4489 "Loop weight_value≤target_weight and delta≟0.0 or delta≥0.01" "noBreak"
        thread Thread_while_4489():
          while (True):
            $ 4490 "MoveL" "noBreak"
            $ 4491 "dispense_pos" "noBreak"
            movel(dispense_pos, a=0.2, v=0.1)
            $ 4492 "prev_weight≔get_weight()" "noBreak"
            global prev_weight=get_weight()
            $ 4493 "log_weight()" "noBreak"
            log_weight()
            $ 4494 "Wait: 0.5" "noBreak"
            sleep(0.5)
            $ 4495 "tilt_pose≔pose_trans(get_actual_tcp_pose(), p[0, 0, 0, 0, 0, 2.0])" "noBreak"
            global tilt_pose=pose_trans(get_actual_tcp_pose(), p[0, 0, 0, 0, 0, 2.0])
            $ 4496 "movel(tilt_pose, a=0.5, v=0.5, r=0.00001)" "noBreak"
            movel(tilt_pose, a=0.5, v=0.5, r=0.00001)
            $ 4497 "weight_value≔get_weight()" "noBreak"
            global weight_value=get_weight()
            $ 4498 "tilt_angle≔-1" "noBreak"
            global tilt_angle=-1
            $ 4499 "Wait: 0.5" "noBreak"
            sleep(0.5)
            $ 4500 "dispense_pos" "noBreak"
            movel(dispense_pos, a=1.2, v=0.25)
            $ 4501 "compute_level_percent(W_now, weight_value)" "noBreak"
            compute_level_percent(W_now, weight_value)
            $ 4502 "prev_spat≔spatula" "noBreak"
            global prev_spat=spatula
            $ 4503 "Wait: 0.2" "noBreak"
            sleep(0.2)
            $ 4505 "spatula≔select_spatula(Flowability, level, diff, bulk_density, mouth_d)" "noBreak"
            global spatula=select_spatula(Flowability, level, diff, bulk_density, mouth_d)
            $ 4506 "Wait: 1.0" "noBreak"
            sleep(1.0)
            $ 4507 "send_level_info()" "noBreak"
            send_level_info()
            $ 4508 "send_spatula_info()" "noBreak"
            send_spatula_info()
            $ 4509 "Set AO[0]=0.0" "noBreak"
            set_standard_analog_out(0, 0.0)
            $ 4510 "Wait: 0.5" "noBreak"
            sleep(0.5)
            $ 4511 "swtich spatula" "noBreak"
            $ 4512 "If spatula ≟ 'spatula_M' and switch_spat_M≟ True " "noBreak"
            if (spatula  ==  "spatula_M"  and  switch_spat_M ==   True  ):
              $ 4513 "MoveJ" "noBreak"
              $ 4514 "Spatula_otw" "noBreak"
              movej(get_inverse_kin(Spatula_otw_p, qnear=Spatula_otw_q), a=1.3962634015954636, v=1.0471975511965976)
              $ 4515 "spat_L_up" "noBreak"
              movej(get_inverse_kin(spat_L_up_p, qnear=spat_L_up_q), a=1.3962634015954636, v=1.0471975511965976)
              $ 4516 "MoveL" "noBreak"
              $ 4517 "spat_L_side" "noBreak"
              movel(spat_L_side_p, a=1.2, v=0.25)
              $ 4518 "spat_L_lift" "noBreak"
              movel(spat_L_lift_p, a=1.2, v=0.25)
              $ 4519 "spat_L_pick" "noBreak"
              movel(spat_L_pick_p, a=0.2, v=0.1)
              # begin: URCap Program Node
              #   Source: Robotiq_Grippers, 3.17.0.105337, Robotiq Inc.
              #   Type: Gripper
              $ 4520 "Gripper Open (1)" "noBreak"
              if not(gripper_connected[0]):
                popup("Gripper 1 must be connected to run this program.", "No connection", False, True, True)
              end
              if not(rq_is_gripper_activated("1")):
                popup("Gripper 1 is not activated. Go to Installation tab > Gripper to activate it and run the program again.", "Not activated", False, True, True)
              end
              rq_set_pos_spd_for(0, 255, 77, "1")
              rq_wait_pos_spe_for_request(0, 255, 77, "1")
              rq_go_to("1")
              rq_wait("1")
              # end: URCap Program Node
              $ 4521 "spat_M_pick" "noBreak"
              movel(spat_M_pick_p, a=1.2, v=0.25)
              # begin: URCap Program Node
              #   Source: Robotiq_Grippers, 3.17.0.105337, Robotiq Inc.
              #   Type: Gripper
              $ 4522 "Gripper Close (1)" "noBreak"
              if not(gripper_connected[0]):
                popup("Gripper 1 must be connected to run this program.", "No connection", False, True, True)
              end
              if not(rq_is_gripper_activated("1")):
                popup("Gripper 1 is not activated. Go to Installation tab > Gripper to activate it and run the program again.", "Not activated", False, True, True)
              end
              rq_set_pos_spd_for(255, 0, 77, "1")
              rq_wait_pos_spe_for_request(255, 0, 77, "1")
              rq_go_to("1")
              rq_wait("1")
              # end: URCap Program Node
              $ 4523 "spat_M_up" "noBreak"
              movel(spat_M_up_p, a=1.2, v=0.25)
              $ 4524 "Spatula_otw" "noBreak"
              movel(Spatula_otw_p, a=1.2, v=0.25)
              $ 4525 "switch_spat_M≔ False " "noBreak"
              global switch_spat_M=  False
              $ 4526 "correction_reset()" "noBreak"
              correction_reset()
            else:
              $ 4527 "ElseIf spatula ≟ 'spatula_S' and switch_spat_S ≟ True and prev_spat≟'spatula_M'" "noBreak"
              if (spatula  ==  "spatula_S" and switch_spat_S  ==   True  and prev_spat == "spatula_M"):
                $ 4528 "MoveL" "noBreak"
                $ 4529 "Spatula_otw" "noBreak"
                movel(Spatula_otw_p, a=1.2, v=0.25)
                $ 4530 "spat_M_up" "noBreak"
                movel(spat_M_up_p, a=1.2, v=0.25)
                $ 4531 "spat_M_pick" "noBreak"
                movel(spat_M_pick_p, a=0.2, v=0.1)
                # begin: URCap Program Node
                #   Source: Robotiq_Grippers, 3.17.0.105337, Robotiq Inc.
                #   Type: Gripper
                $ 4532 "Gripper Open (1)" "noBreak"
                if not(gripper_connected[0]):
                  popup("Gripper 1 must be connected to run this program.", "No connection", False, True, True)
                end
                if not(rq_is_gripper_activated("1")):
                  popup("Gripper 1 is not activated. Go to Installation tab > Gripper to activate it and run the program again.", "Not activated", False, True, True)
                end
                rq_set_pos_spd_for(0, 255, 77, "1")
                rq_wait_pos_spe_for_request(0, 255, 77, "1")
                rq_go_to("1")
                rq_wait("1")
                # end: URCap Program Node
                $ 4533 "spat_S_pick" "noBreak"
                movel(spat_S_pick_p, a=1.2, v=0.25)
                # begin: URCap Program Node
                #   Source: Robotiq_Grippers, 3.17.0.105337, Robotiq Inc.
                #   Type: Gripper
                $ 4534 "Gripper Close (1)" "noBreak"
                if not(gripper_connected[0]):
                  popup("Gripper 1 must be connected to run this program.", "No connection", False, True, True)
                end
                if not(rq_is_gripper_activated("1")):
                  popup("Gripper 1 is not activated. Go to Installation tab > Gripper to activate it and run the program again.", "Not activated", False, True, True)
                end
                rq_set_pos_spd_for(255, 0, 77, "1")
                rq_wait_pos_spe_for_request(255, 0, 77, "1")
                rq_go_to("1")
                rq_wait("1")
                # end: URCap Program Node
                $ 4535 "spat_S_up" "noBreak"
                movel(spat_S_up_p, a=1.2, v=0.25)
                $ 4536 "Spatula_otw" "noBreak"
                movel(Spatula_otw_p, a=1.2, v=0.25)
                $ 4537 "switch_spat_S≔ False " "noBreak"
                global switch_spat_S=  False
                $ 4538 "correction_reset()" "noBreak"
                correction_reset()
              else:
                $ 4539 "ElseIf spatula≟'spatula_S' and switch_spat_S≟ True  and prev_spat≟'spatula_L'" "noBreak"
                if (spatula == "spatula_S" and switch_spat_S ==   True    and  prev_spat == "spatula_L"):
                  $ 4540 "MoveJ" "noBreak"
                  $ 4541 "Spatula_otw" "noBreak"
                  movej(get_inverse_kin(Spatula_otw_p, qnear=Spatula_otw_q), a=1.3962634015954636, v=1.0471975511965976)
                  $ 4542 "spat_L_up" "noBreak"
                  movej(get_inverse_kin(spat_L_up_p, qnear=spat_L_up_q), a=1.3962634015954636, v=1.0471975511965976)
                  $ 4543 "MoveL" "noBreak"
                  $ 4544 "spat_L_side" "noBreak"
                  movel(spat_L_side_p, a=1.2, v=0.25)
                  $ 4545 "spat_L_lift" "noBreak"
                  movel(spat_L_lift_p, a=1.2, v=0.25)
                  $ 4546 "spat_L_pick" "noBreak"
                  movel(spat_L_pick_p, a=0.2, v=0.1)
                  # begin: URCap Program Node
                  #   Source: Robotiq_Grippers, 3.17.0.105337, Robotiq Inc.
                  #   Type: Gripper
                  $ 4547 "Gripper Open (1)" "noBreak"
                  if not(gripper_connected[0]):
                    popup("Gripper 1 must be connected to run this program.", "No connection", False, True, True)
                  end
                  if not(rq_is_gripper_activated("1")):
                    popup("Gripper 1 is not activated. Go to Installation tab > Gripper to activate it and run the program again.", "Not activated", False, True, True)
                  end
                  rq_set_pos_spd_for(0, 255, 77, "1")
                  rq_wait_pos_spe_for_request(0, 255, 77, "1")
                  rq_go_to("1")
                  rq_wait("1")
                  # end: URCap Program Node
                  $ 4548 "spat_S_pick" "noBreak"
                  movel(spat_S_pick_p, a=1.2, v=0.25)
                  # begin: URCap Program Node
                  #   Source: Robotiq_Grippers, 3.17.0.105337, Robotiq Inc.
                  #   Type: Gripper
                  $ 4549 "Gripper Close (1)" "noBreak"
                  if not(gripper_connected[0]):
                    popup("Gripper 1 must be connected to run this program.", "No connection", False, True, True)
                  end
                  if not(rq_is_gripper_activated("1")):
                    popup("Gripper 1 is not activated. Go to Installation tab > Gripper to activate it and run the program again.", "Not activated", False, True, True)
                  end
                  rq_set_pos_spd_for(255, 0, 77, "1")
                  rq_wait_pos_spe_for_request(255, 0, 77, "1")
                  rq_go_to("1")
                  rq_wait("1")
                  # end: URCap Program Node
                  $ 4550 "spat_S_up" "noBreak"
                  movel(spat_S_up_p, a=1.2, v=0.25)
                  $ 4551 "Spatula_otw" "noBreak"
                  movel(Spatula_otw_p, a=1.2, v=0.25)
                  $ 4552 "switch_spat_S≔ False " "noBreak"
                  global switch_spat_S=  False
                  $ 4553 "correction_reset()" "noBreak"
                  correction_reset()
                else:
                  $ 4554 "ElseIf spatula≟'spatula_flat_S'  and switch_spat_F_S ≟ True " "noBreak"
                  if (spatula == "spatula_flat_S"   and  switch_spat_F_S  ==   True  ):
                    $ 4555 "MoveL" "noBreak"
                    $ 4556 "Spatula_otw" "noBreak"
                    movel(Spatula_otw_p, a=1.2, v=0.25)
                    $ 4557 "spat_flatM_up" "noBreak"
                    movel(spat_flatM_up_p, a=1.2, v=0.25)
                    $ 4558 "spat_flatM_pick" "noBreak"
                    movel(spat_flatM_pick_p, a=0.2, v=0.1)
                    # begin: URCap Program Node
                    #   Source: Robotiq_Grippers, 3.17.0.105337, Robotiq Inc.
                    #   Type: Gripper
                    $ 4559 "Gripper Open (1)" "noBreak"
                    if not(gripper_connected[0]):
                      popup("Gripper 1 must be connected to run this program.", "No connection", False, True, True)
                    end
                    if not(rq_is_gripper_activated("1")):
                      popup("Gripper 1 is not activated. Go to Installation tab > Gripper to activate it and run the program again.", "Not activated", False, True, True)
                    end
                    rq_set_pos_spd_for(0, 0, 77, "1")
                    rq_wait_pos_spe_for_request(0, 0, 77, "1")
                    rq_go_to("1")
                    rq_wait("1")
                    # end: URCap Program Node
                    $ 4560 "spat_flatS_pick" "noBreak"
                    movel(spat_flatS_pick_p, a=1.2, v=0.25)
                    # begin: URCap Program Node
                    #   Source: Robotiq_Grippers, 3.17.0.105337, Robotiq Inc.
                    #   Type: Gripper
                    $ 4561 "Gripper Close (1)" "noBreak"
                    if not(gripper_connected[0]):
                      popup("Gripper 1 must be connected to run this program.", "No connection", False, True, True)
                    end
                    if not(rq_is_gripper_activated("1")):
                      popup("Gripper 1 is not activated. Go to Installation tab > Gripper to activate it and run the program again.", "Not activated", False, True, True)
                    end
                    rq_set_pos_spd_for(255, 0, 77, "1")
                    rq_wait_pos_spe_for_request(255, 0, 77, "1")
                    rq_go_to("1")
                    rq_wait("1")
                    # end: URCap Program Node
                    $ 4562 "spat_flatS_up" "noBreak"
                    movel(spat_flatS_up_p, a=1.2, v=0.25)
                    $ 4563 "Spatula_otw" "noBreak"
                    movel(Spatula_otw_p, a=1.2, v=0.25)
                    $ 4564 "switch_spat_F_S≔ False " "noBreak"
                    global switch_spat_F_S=  False
                    $ 4565 "correction_reset()" "noBreak"
                    correction_reset()
                  end
                end
              end
            end
            $ 4566 "tilt(level)" "noBreak"
            tilt(level)
            $ 4567 "Action_Info≔'Scooping'" "noBreak"
            global Action_Info="Scooping"
            $ 4568 "auto_tilt_and_scoop(W_now, target_weight, weight_value)" "noBreak"
            auto_tilt_and_scoop(W_now, target_weight, weight_value)
            $ 4569 "Action_Info≔'Dosing'" "noBreak"
            global Action_Info="Dosing"
          end
        end
        if (weight_value <= target_weight and delta == 0.0 or delta >= 0.01):
          global thread_handler_4489=run Thread_while_4489()
